(* CODESYS project lc.library
   DefaultNamespace: KOSTAL.AF2024.Connectivity.LC
   DocFormat: reStructuredText
   Description: Contains Components to communicate with LC Webservice.
      
      Designed with webAPI Version 2.0.39
      
      =====================
      BASED NOT ON I_LC!!
      =====================
   Author: Frank Dümpelmann
   Title: KOSTAL.AF2024.Connectivity.LC
   Version: 1.0.0.0
   Company: KOSTAL GmbH & Co.KG
   Placeholder: KOSTAL.AF2024.Connectivity.LC

Project tree, tasks and I/O mapping:
  libraries: KOSTAL.AF2024.Connectivity.TLS.CipherSuite.OpenSSL, 1.0.0.0 (KOSTAL GmbH & Co.KG); KOSTAL.AF2024.Core.FileLogger, 1.0.0.0 (KOSTAL GmbH & Co.KG); KOSTAL.AF2024.Core.functionResponse, 1.0.0.0 (KOSTAL GmbH & Co.KG); KOSTAL.AF2024.Core.GetSystemTime, 1.0.1.0 (KOSTAL GmbH & Co.KG); KOSTAL.AF2024.Core.JsonTools, 1.0.0.0 (KOSTAL GmbH & Co.KG); KOSTAL.AF2024.Core.ListOf, 1.0.0.0 (KOSTAL GmbH & Co.KG); KOSTAL.AF2024.Core.Process, 1.0.1.0 (KOSTAL GmbH & Co.KG); KOSTAL.AF2024.Core.Settings, 1.0.0.0 (KOSTAL GmbH & Co.KG); KOSTAL.AF2024.Core.StringTools, 1.0.0.0 (KOSTAL GmbH & Co.KG); KOSTAL.AF2024.Core.System, 1.0.0.0 (KOSTAL GmbH & Co.KG); Tc2_Standard, 3.4.5.0 (Beckhoff Automation GmbH); Tc2_System, 3.6.4.0 (Beckhoff Automation GmbH); Tc2_Utilities, 3.7.4.0 (Beckhoff Automation GmbH); Tc3_IotBase, 3.4.5.0 (Beckhoff Automation GmbH); Tc3_JsonXml, 3.4.4.0 (Beckhoff Automation GmbH)
  0_Internal/
    interface _I_T_Copy: CopyTo
    interface _I_T_Copy_Owner: Clear, CopyFrom, CopyTo
    interface _I_T_CopyFrom: CopyFrom
    function block _T_Copy [ST]: Clear, CopyFrom, CopyTo
  1_Config/
    Reader/
      DUT/
        interface I_T_Header: CopyTo, ID, name, sourceName, timeStamp
        interface I_T_Header_CopyFrom: CopyFrom
        function block T_Header [ST]: Clear, CopyFrom, CopyTo, ID, name, sourceName, timeStamp
      function block FB_Reader [ST]: _Step_ClearContent, _Step_ParseContent, CFG, Header
      global variables JSON_MEMBER
    interface I_T_CFG: ClientName, ClientProcess, CopyTo, HostName, HostPort, Valid
    interface I_T_CFG_CopyFrom: CopyFrom
    function block T_CFG [ST]: Clear, ClientName, ClientProcess, CopyFrom, CopyTo, HostName, HostPort, Valid
  2_BaseClass/
    DUT/
      Response/
        interface I_T_ResponseResult: CopyTo, errorMessage, internalDuration, isErrorOccured, isResultGood
        interface I_T_ResponseResult_CopyFrom: CopyFrom
        interface I_T_ResponseResult_Owner: clear, CopyFrom, CopyTo, errorMessage, internalDuration, isErrorOccured, isResultGood
        function block T_ResponseResult [ST]: clear, CopyFrom, CopyTo, errorMessage, internalDuration, isErrorOccured, isResultGood
      data type E_PROCESS
      data type E_Verbose
    POE/
      function block FB_LC [ST]: _getResponseResultFromJson, _PARSE_ARRAY, _PARSE_BOOL, _PARSE_BYTE, _PARSE_DINT, _PARSE_JSON, _PARSE_STRING, _PARSE_TIME, _PARSE_UDINT, _PARSE_ULINT, _00_clientCfg, _01_Ready, _10_finishFail, _10_finishPass, _10_GET, _10_GET_CTRL, _10_GET_ResponseResult, _10_GET_ResponseResult_CTRL, _10_SET, _10_SET_CTRL, _99_stepError, _CfgChange, _CfgHasChanged, _deviceDefine, _logStartMessage, _UriGet, _UrlReplace, _VerboseHandler, ClientName, ClientProcess, HostName, HostPort, HTTP_Statuscode, IN_PROCESS, KeepAlive, repeatsOnFail, State, TimeOut, WS_Duration, FBmain, GetTimeStamp, linkConfig, LinkTime, RedirectClient, Verbose, _FBmain
  3_DUT/
    OptionalFlags/
      interface I_T_OptionalFlags: FlagsInRange, get
      interface I_T_OptionalFlags_Owner: clear, FlagsInRange, get, set
      function block T_OptionalFlags [ST]: clear, CopyFrom, FlagsInRange, get, set
    OptionalStrings/
      interface I_T_OptionalStrings: get, StringsInRange
      interface I_T_OptionalStrings_Owner: clear, get, set, StringsInRange
      function block T_OptionalStrings [ST]: clear, CopyFrom, get, set, StringsInRange
    PreviousProcess/
      ListOf/
        function block FB_ListOfPreviousProcess [ST]: _get_I, _get_I_Owner, _removePayLoad, _verifyMember, Add_DUT, Clear, CopyFrom, CopyTo, Delete_DUT, Get_I, Get_I_ByProcessName, Get_I_Owner, NumberOfMember
        interface I_ListOfPreviousProcess: CopyTo, Get_I, Get_I_ByProcessName, NumberOfMember
        interface I_ListOfPreviousProcess_CopyFrom: CopyFrom
        interface I_ListOfPreviousProcess_Owner: Add_DUT, Clear, CopyFrom, CopyTo, Delete_DUT, Get_I, Get_I_ByProcessName, Get_I_Owner, NumberOfMember
      interface I_T_PreviousProcess: articlenumberRegex, databaseName, PreviousProcesses, processName, processStamp, searchMode, useOnlyTable
      interface I_T_PreviousProcess_Owner: articlenumberRegex, clear, databaseName, PreviousProcesses_Owner, processName, processStamp, searchMode, useOnlyTable
      function block T_PreviousProcess [ST]: articlenumberRegex, clear, CopyFrom, databaseName, PreviousProcesses, PreviousProcesses_Owner, processName, processStamp, searchMode, useOnlyTable
    ProcessConfig/
      ListOf/
        function block FB_ListOfProcessConfig [ST]: _get_I, _get_I_Owner, _removePayLoad, _verifyMember, Add_DUT, Clear, CopyFrom, CopyTo, Delete_DUT, Get_I, Get_I_Owner, NumberOfMember
        interface I_ListOfProcessConfig: CopyTo, Get_I, NumberOfMember
        interface I_ListOfProcessConfig_CopyFrom: CopyFrom
        interface I_ListOfProcessConfig_Owner: Add_DUT, Clear, CopyFrom, CopyTo, Delete_DUT, Get_I, Get_I_Owner, NumberOfMember
      interface I_T_ProcessConfig: activeCheckFQDN, allowedFQDN, articlenumberRegex, PreviousProcesses, serialnumberRegex, traceID
      interface I_T_ProcessConfig_Owner: activeCheckFQDN, allowedFQDN, articlenumberRegex, clear, PreviousProcesses_Owner, serialnumberRegex, traceID
      function block T_ProcessConfig [ST]: activeCheckFQDN, allowedFQDN, articlenumberRegex, clear, CopyFrom, PreviousProcesses, PreviousProcesses_Owner, serialnumberRegex, traceID
    SingleProcess/
      ListOf/
        function block FB_ListOfSingleProcess [ST]: _get_I, _get_I_Owner, _removePayLoad, _verifyMember, Add_DUT, Clear, CopyFrom, CopyTo, Delete_DUT, Get_I, Get_I_Owner, NumberOfMember
        interface I_ListOfSingleProcess: CopyTo, Get_I, NumberOfMember
        interface I_ListOfSingleProcess_CopyFrom: CopyFrom
        interface I_ListOfSingleProcess_Owner: Add_DUT, Clear, CopyFrom, CopyTo, Delete_DUT, Get_I, Get_I_Owner, NumberOfMember
      interface I_T_SingleProcess: articleNumber, id, OptionalFlags, OptionalStrings, process, result, serialNumber, timeStamp, traceId
      interface I_T_SingleProcess_Owner: articleNumber, clear, id, OptionalFlags_Owner, OptionalStrings_Owner, process, result, serialNumber, timeStamp, traceId
      function block T_SingleProcess [ST]: articleNumber, clear, CopyFrom, id, OptionalFlags, OptionalFlags_Owner, OptionalStrings, OptionalStrings_Owner, process, result, serialNumber, timeStamp, traceId
    SubModule/
      ListOf/
        function block FB_ListOfSubModule [ST]: _get_I, _get_I_Owner, _removePayLoad, _verifyMember, Add_DUT, Clear, CopyFrom, CopyTo, Delete_DUT, Get_I, Get_I_Owner, NumberOfMember
        interface I_ListOfSubModule: CopyTo, Get_I, NumberOfMember
        interface I_ListOfSubModule_CopyFrom: CopyFrom
        interface I_ListOfSubModule_Owner: Add_DUT, Clear, CopyFrom, CopyTo, Delete_DUT, Get_I, Get_I_Owner, NumberOfMember
      interface I_T_SubModule: articleNumber, serialNumber
      interface I_T_SubModule_Owner: articleNumber, clear, serialNumber
      function block T_SubModule [ST]: articleNumber, clear, CopyFrom, serialNumber
    SubModuleOfProcess/
      ListOf/
        function block FB_ListOfSubModuleOfProcess [ST]: _get_I, _get_I_Owner, _removePayLoad, _verifyMember, Add_DUT, Clear, CopyFrom, CopyTo, Delete_DUT, Get_I, Get_I_Owner, NumberOfMember
        interface I_ListOfSubModuleOfProcess: CopyTo, Get_I, NumberOfMember
        interface I_ListOfSubModuleOfProcess_CopyFrom: CopyFrom
        interface I_ListOfSubModuleOfProcess_Owner: Add_DUT, Clear, CopyFrom, CopyTo, Delete_DUT, Get_I, Get_I_Owner, NumberOfMember
      interface I_T_SubModuleOfProcess: timeStamp
      interface I_T_SubModuleOfProcess_Owner: timeStamp
      function block T_SubModuleOfProcess [ST]: clear, CopyFrom, timeStamp
    WriteCurrentStampDataDto/
      interface I_T_WriteCurrentStampDataDto: articleNumber, OptionalFlags, OptionalStrings, result, serialNumber
      interface I_T_WriteCurrentStampDataDto_Owner: articleNumber, clear, OptionalFlags_Owner, OptionalStrings_Owner, result, serialNumber
      function block T_WriteCurrentStampDataDto [ST]: articleNumber, clear, CopyFrom, OptionalFlags, OptionalFlags_Owner, OptionalStrings, OptionalStrings_Owner, result, serialNumber
  4_GVL/
    global variables API_VERSION
    global variables PROCESS_CONFIG
    global variables PROCESS_INFO
    global variables RESPONSE_BODY
    global variables SETTINGS
    global variables SUBMODUL_INFO
    global variables URL
  5_POU/
    GetetParentBySubmoduleSerialnumber/
      function block FB_GetParent_By_SM_SN [ST]: _getProcessInfo, _getSubModule_n, _getSubModuleList, _01_Ready, _10_getProcessInfo, _10_getSubModule_n, _10_getSubModuleList, _10_processRead, _selectUrl, Execute, ListOfSubModules, ResponseProcess, ResponseResult, _FBmain
    GetSubModulesByParentSerialNumber/
      function block FB_GetSM_ByParentSN [ST]: _getProcessInfo, _getSubModule_n, _getSubModuleList, _01_Ready, _10_getProcessInfo, _10_getSubModule_n, _10_getSubModuleList, _10_processRead, _selectUrl, Execute, ListOfSubModules, ResponseProcess, ResponseResult, _FBmain
    Init/
      function block FB_Init [ST]
    ReadApiVersion/
      MustBeExtended/
        function block _FB_ReadApiVersion [ST]: _getApiVersion, _01_Ready, _10_getapiVersion, _10_processRead, _selectUrl, apiVersion, ResponseResult, _FBmain
      function block FB_ReadApiVersion [ST]: Execute, _selectUrl
    ReadProcess/
      MustBeExtended/
        function block _FB_ReadProcess [ST]: _getProcessInfo, _getProcessInfoList, _01_Ready, _10_getProcessInfo_n, _10_getProcessInfoList, _10_processRead, _selectUrl, GetSingleProcess, NumberOfSingleProcess, ProcessInfoListLenght, ResponseResult, _FBmain
      function block FB_ReadPreviousProcess_SN [ST]: Execute, _selectUrl
      function block FB_ReadPreviousProcess_SN_ART [ST]: Execute, _selectUrl
      function block FB_ReadProcess_ID [ST]: Execute, _selectUrl
      function block FB_ReadProcess_SN [ST]: Execute, _selectUrl
      function block FB_ReadProcess_SN_ART [ST]: Execute, _selectUrl
    ReadProcessConfig/
      MustBeExtended/
        function block _FB_ReadConfig [ST]: _getPreviousProcess, _getPreviousProcesses, _getPreviousProcessList, _getProcessConfig, _getProcessConfigList, _01_Ready, _10_getProcessConfig_n, _10_getProcessConfigList, _10_processRead, _selectUrl, GetProcessConfig, NumberOfProcessConfig, ResponseResult, _FBmain
      function block FB_ReadProcessConfig [ST]: Execute, _selectUrl
    WriteProcess/
      MustBeExtended/
        function block _FB_WriteProcess [ST]: _getProcessInfo, _01_Ready, _10_getProcessInfo, _10_processWrite, _20_setProcessInfo, _selectUrl, Execute, ResponseProcess, ResponseResult, WriteDataDto
      function block FB_WriteProcess [ST]: _selectUrl, _FBmain
      function block FB_WriteProcessWithSM [ST]: _20_setSubModules, _selectUrl, ListOfSubModules, _FBmain
  Project Information/
    function F_GetCompany [ST]
    function F_GetTitle [ST]
    function F_GetVersion [ST]
  Version/
    global variables Global_Version
*)

// 2_BaseClass/DUT/E_PROCESS
{attribute 'qualified_only'}
{attribute 'strict'}
TYPE E_PROCESS :
(
	idle		:= 0,
	execute	:= 1
);
END_TYPE

// 2_BaseClass/DUT/E_Verbose
{attribute 'qualified_only'}
{attribute 'strict'}
(*
Note that the verbose status is evaluated binary
================================================
*)
TYPE E_Verbose :
(
	none 			:= 0,
	Request		:= 1,
	Response	:= 2,
	Both			:= 3
);
END_TYPE

// 1_Config/Reader/JSON_MEMBER
{attribute 'qualified_only'}
VAR_GLOBAL CONSTANT

	{region 'Header'}
		ID					: STRING:= 'ID';
		name				: STRING:= 'name'; 
		timeStamp		: STRING:= 'timeStamp'; 
		sourceName	: STRING:= 'sourceName'; 
	{endregion}

	{region 'LC'}
		LC						: STRING:= 'LC';
		HostName			: STRING:= 'HostName';
		HostPort			: STRING:= 'HostPort';
		ClientName		: STRING:= 'ClientName';
		ClientProcess	: STRING:= 'ClientProcess';
	{endregion}

END_VAR

// 4_GVL/API_VERSION
{attribute 'qualified_only'}
VAR_GLOBAL
	apiVersion		:	STRING:= 'apiVersion';
END_VAR

// 4_GVL/PROCESS_CONFIG
{attribute 'qualified_only'}
VAR_GLOBAL CONSTANT
	//
	processConfiguration	:	STRING:=	'processConfiguration';
	//
  articlenumberRegex	: STRING:=	'articlenumberRegex';	//"^[0-9]{8}-(([0-9]{2})|([0-9]{4}))$",
  serialnumberRegex		: STRING:=	'serialnumberRegex';	//"^([A-Z0-9]{13})$|^([0-9]{14})$",
  traceID							: STRING:=	'traceID';	//99056,
	activeCheckFQDN			: STRING:=	'activeCheckFQDN';
	allowedFQDN					: STRING:=	'allowedFQDN';
	///--
  previousProcesses	: STRING:=	'previousProcesses';	//[...]
	//
  processName			: STRING:=	'processName';	//"ASS01",
  processStamp		: STRING:=	'processStamp';	//"ASS01",
  databaseName		: STRING:=	'databaseName';		//"test",
  useOnlyTable		: STRING:=	'useOnlyTable';	//"lc_test"
  searchMode			: STRING:=	'searchMode';	//0,
  //articlenumberRegex	: STRING:=	'articlenumberRegex';	same as in parent node
  //previousProcesses	: STRING:=	'previousProcesses';	same as in parent node

//obsolete
//  databaseServer	:	STRING:=	'databaseServer';	//"debelc034.de.kostal.int",
//  databasePort		: STRING:=	'databasePort';		//3306,
//  databaseUser		: STRING:=	'databaseUser';		//null,
END_VAR

// 4_GVL/PROCESS_INFO
{attribute 'qualified_only'}
VAR_GLOBAL CONSTANT
	//
	processInfoList	: STRING:= 'processInfoList'; 
	processInfo			: STRING:= 'processInfo';
	//
	id								: STRING:= 'id';
	serialNumber			: STRING:= 'serialNumber';
	articleNumber			: STRING:= 'articleNumber';
	timeStamp					: STRING:= 'timeStamp';
	traceId						: STRING:= 'traceId';
	process						: STRING:= 'process';
	result						: STRING:= 'result';
	optionalString_1	: STRING:= 'optionalString_1';
	optionalString_2	: STRING:= 'optionalString_2';
	optionalString_3	: STRING:= 'optionalString_3';
	optionalString_4	: STRING:= 'optionalString_4';
	optionalFlag_1		: STRING:= 'optionalFlag_1';
	optionalFlag_2		: STRING:= 'optionalFlag_2';
	optionalFlag_3		: STRING:= 'optionalFlag_3';
	optionalFlag_4		: STRING:= 'optionalFlag_4';
	optionalFlag_5		: STRING:= 'optionalFlag_5';
	optionalFlag_6		: STRING:= 'optionalFlag_6';
	optionalFlag_7		: STRING:= 'optionalFlag_7';
	optionalFlag_8		: STRING:= 'optionalFlag_8';

	//
	childs	: STRING:= 'Childs';
																		
END_VAR

// 4_GVL/RESPONSE_BODY
{attribute 'qualified_only'}
VAR_GLOBAL CONSTANT
	
	isErrorOccured		:	STRING:= 'isErrorOccured';
	isResultGood			:	STRING:= 'isResultGood';
	errorMessage			:	STRING:= 'errorMessage';
	internalDuration	:	STRING:= 'internalDuration';
	
END_VAR

// 4_GVL/SETTINGS
{attribute 'qualified_only'}
VAR_GLOBAL CONSTANT
	OPTIONAL_FLAGS_MAX				: UINT:= 8;
	
	OPTIONAL_STRINGS_MAX			: UINT:= 4;
	OPTIONAL_STRINGS_LENGHT		: UINT:= SIZEOF(KOSTAL_AF2024_Core_Settings.T_MaxString_UTF8);
END_VAR

// 4_GVL/SUBMODUL_INFO
{attribute 'qualified_only'}
VAR_GLOBAL CONSTANT
	//
	subModules	: STRING:= 'submodules';
	//
	serialNumber	: STRING:=	'serialNumber';
	articleNumber : STRING:=	'articleNumber';
	timestamp			: STRING:=	'timestamp';	//only in S´sub modules of process available
END_VAR

// 4_GVL/URL
{attribute 'qualified_only'}
VAR_GLOBAL CONSTANT

	URI_BASE	: KOSTAL_AF2024_Core_Settings.T_MaxString_UTF8:=  '/ws/api/gen2/';
	
	READ_API_VERSION	: KOSTAL_AF2024_Core_Settings.T_MaxString_UTF8:= 'readApiVersion';
	
	READ_PROC_RECORD_ID	: KOSTAL_AF2024_Core_Settings.T_MaxString_UTF8:= 'readProcess/{ClientName}/{ClientProcess}/id={RecordID}';

	READ_PROC_SERNO				: KOSTAL_AF2024_Core_Settings.T_MaxString_UTF8:= 'readProcess/{ClientName}/{ClientProcess}/{SerialNumber}';
	READ_PROCESS_SERNO_OPT_PROC	: KOSTAL_AF2024_Core_Settings.T_MaxString_UTF8:= 'readProcess/{ClientName}/{ClientProcess}/{SerialNumber}?Process={?Process=}';
	
	READ_PROC_SERNO_ARTNO			: KOSTAL_AF2024_Core_Settings.T_MaxString_UTF8:= 'readProcess/{ClientName}/{ClientProcess}/{SerialNumber}/{ArticleNumber}';
	READ_PROC_SERNO_ARTNO_OPT_PROC	: KOSTAL_AF2024_Core_Settings.T_MaxString_UTF8:= 'readProcess/{ClientName}/{ClientProcess}/{SerialNumber}/{ArticleNumber}?Process={?Process=}';

	READ_PREV_PROC_SERNO	: KOSTAL_AF2024_Core_Settings.T_MaxString_UTF8:= 'readPreviousProcess/{ClientName}/{ClientProcess}/{SerialNumber}';

	READ_PREV_PROC_SERNO_ARTNO	: KOSTAL_AF2024_Core_Settings.T_MaxString_UTF8:= 'readPreviousProcess/{ClientName}/{ClientProcess}/{SerialNumber}/{ArticleNumber}';
	
	WRITE_CUR_PROC					: KOSTAL_AF2024_Core_Settings.T_MaxString_UTF8:= 'writeCurrentProcess/{ClientName}/{ClientProcess}';
	WRITE_CUR_PROC_WITH_SUBMODULS	: KOSTAL_AF2024_Core_Settings.T_MaxString_UTF8:= 'writeCurrentProcessWithSubmodules/{ClientName}/{ClientProcess}';

	READ_PROC_CONF			: KOSTAL_AF2024_Core_Settings.T_MaxString_UTF8:= 'readProcessConfig/{ClientName}';
	READ_PROC_CONF_OPT_PROC	: KOSTAL_AF2024_Core_Settings.T_MaxString_UTF8:= 'readProcessConfig/{ClientName}/{ClientProcess}';

	READ_SUB_MODULES_BY_PARENT_SERIAL_NUMBER	: KOSTAL_AF2024_Core_Settings.T_MaxString_UTF8:= 'getSubmodulesByParentserialnumber/{ClientName}/{ClientProcess}/{ParentSerialnumber}';
	READ_PARENT_BY_SUB_MODULE_SERIAL_NUMBER		: KOSTAL_AF2024_Core_Settings.T_MaxString_UTF8:= 'getParentBySubmoduleSerialnumber/{ClientName}/{ClientProcess}/{SubmoduleSerialnumber}';
END_VAR

//Placeholder for URI
{attribute 'qualified_only'}
VAR_GLOBAL CONSTANT
	PLACEHOLDER_CLIENT_NAME						: STRING:= '{ClientName}';
	PLACEHOLDER_CLIENT_PROCESS				: STRING:= '{ClientProcess}';
	PLACEHOLDER_RECORD_ID							: STRING:= '{RecordID}';
	PLACEHOLDER_SERIALNUMBER					: STRING:= '{SerialNumber}';
	PLACEHOLDER_ARTICLENUMBER					: STRING:= '{ArticleNumber}';
	PLACEHOLDER_OPTIONAL_PROCESS			: STRING:= '{?Process=}';

	PLACEHOLDER_PARENT_SERIAL_NUMBER	: STRING:= '{ParentSerialnumber}';
	PLACEHOLDER_SUB_MODULE_SERIAL_NUMBER		: STRING:= '{SubmoduleSerialnumber}';
END_VAR

// Version/Global_Version
{attribute 'TcGenerated'}
{attribute 'no-analysis'}
{attribute 'linkalways'}
// This function has been automatically generated from the project information.
VAR_GLOBAL CONSTANT
	{attribute 'const_non_replaced'}
	stLibVersion_KOSTAL_AF2024_Connectivity_LC : ST_LibVersion := (iMajor := 1, iMinor := 0, iBuild := 0, iRevision := 0, nFlags := 1, sVersion := '1.0.0.0');
END_VAR

// 0_Internal/_I_T_Copy
INTERFACE _I_T_Copy EXTENDS KOSTAL_AF2024_Core_System.I_Interface

METHOD PUBLIC CopyTo : BOOL
VAR_INPUT
	IN	: KOSTAL_AF2024_Core_System.I_Interface;
END_VAR
END_METHOD

END_INTERFACE

// 0_Internal/_I_T_Copy_Owner
INTERFACE _I_T_Copy_Owner EXTENDS KOSTAL_AF2024_Core_System.I_Interface

METHOD PUBLIC Clear
END_METHOD

METHOD PUBLIC CopyFrom : BOOL
VAR_INPUT
	IN	: KOSTAL_AF2024_Core_System.I_Interface;
END_VAR
END_METHOD

METHOD PUBLIC CopyTo : BOOL
VAR_INPUT
	IN	: KOSTAL_AF2024_Core_System.I_Interface;
END_VAR
END_METHOD

END_INTERFACE

// 0_Internal/_I_T_CopyFrom
INTERFACE _I_T_CopyFrom EXTENDS KOSTAL_AF2024_Core_System.I_Interface

METHOD PUBLIC CopyFrom : BOOL
VAR_INPUT
	IN	: KOSTAL_AF2024_Core_System.I_Interface;
END_VAR
END_METHOD

END_INTERFACE

// 0_Internal/_T_Copy
FUNCTION_BLOCK ABSTRACT _T_Copy IMPLEMENTS _I_T_Copy, _I_T_Copy_Owner, _I_T_CopyFrom

METHOD PUBLIC Clear
END_METHOD

METHOD PUBLIC CopyFrom : BOOL
VAR_INPUT
	IN	: KOSTAL_AF2024_Core_System.I_Interface;
END_VAR

VAR
	_IN	: KOSTAL_AF2024_Core_System.I_Interface;
END_VAR


CopyFrom:= (IN <> 0) AND_THEN __QUERYINTERFACE(IN, _IN) AND_THEN (_IN <> 0);
END_METHOD

METHOD PUBLIC CopyTo : BOOL
VAR_INPUT
	IN	: KOSTAL_AF2024_Core_System.I_Interface;
END_VAR

VAR
	_IN	: _I_T_CopyFrom;
END_VAR

IF (IN = 0) OR_ELSE NOT __QUERYINTERFACE(IN, _IN) OR_ELSE (_IN = 0) THEN	RETURN;	END_IF

CopyTo:= _IN.CopyFrom(THIS^);
END_METHOD

END_FUNCTION_BLOCK

// 1_Config/Reader/DUT/I_T_Header
INTERFACE I_T_Header EXTENDS KOSTAL_AF2024_Core_System.I_Interface

METHOD PUBLIC CopyTo : BOOL
VAR_INPUT
	IN	: I_T_Header_CopyFrom;
END_VAR
END_METHOD

PROPERTY PUBLIC ID : KOSTAL_AF2024_Core_Settings.T_MaxString_UTF8
GET
END_GET
END_PROPERTY

PROPERTY PUBLIC name : KOSTAL_AF2024_Core_Settings.T_MaxString_UTF8
GET
END_GET
END_PROPERTY

PROPERTY PUBLIC sourceName : KOSTAL_AF2024_Core_Settings.T_MaxString_UTF8
GET
END_GET
END_PROPERTY

PROPERTY PUBLIC timeStamp : KOSTAL_AF2024_Core_Settings.T_MaxString_UTF8
GET
END_GET
END_PROPERTY

END_INTERFACE

// 1_Config/Reader/DUT/I_T_Header_CopyFrom
INTERFACE I_T_Header_CopyFrom EXTENDS KOSTAL_AF2024_Core_System.I_Interface

METHOD PUBLIC CopyFrom
VAR_INPUT
	IN	: KOSTAL_AF2024_Core_System.I_Interface;
END_VAR
END_METHOD

END_INTERFACE

// 1_Config/Reader/DUT/T_Header
FUNCTION_BLOCK PUBLIC T_Header IMPLEMENTS I_T_Header, I_T_Header_CopyFrom

VAR
	_ID					: KOSTAL_AF2024_Core_Settings.T_MaxString_UTF8;
	_name				: KOSTAL_AF2024_Core_Settings.T_MaxString_UTF8;
	_timeStamp	: KOSTAL_AF2024_Core_Settings.T_MaxString_UTF8;
	_sourceName	: KOSTAL_AF2024_Core_Settings.T_MaxString_UTF8;	
END_VAR

METHOD PUBLIC Clear
VAR_INPUT
END_VAR

_ID					:= '';
_name				:= '';
_sourceName	:= '';
_timeStamp	:= '';
END_METHOD

METHOD PUBLIC CopyFrom
VAR_INPUT
	IN	: KOSTAL_AF2024_Core_System.I_Interface;
END_VAR

VAR
	_IN	: I_T_Header;
END_VAR

IF IN = 0 THEN	RETURN;	END_IF
IF NOT __QUERYINTERFACE(IN, _IN) OR_ELSE _IN = 0 THEN RETURN;	END_IF

_ID					:= _IN.ID;
_name				:= _IN.name;
_timeStamp	:= _IN.timeStamp;
_sourceName	:= _IN.sourceName;
END_METHOD

METHOD PUBLIC CopyTo : BOOL
VAR_INPUT
	IN	: I_T_Header_CopyFrom;
END_VAR

IF IN = 0 THEN	RETURN;	END_IF

IN.CopyFrom(THIS^);
END_METHOD

PROPERTY PUBLIC ID : KOSTAL_AF2024_Core_Settings.T_MaxString_UTF8
GET

ID:= _ID;
END_GET
SET

_ID:= ID;
END_SET
END_PROPERTY

PROPERTY PUBLIC name : KOSTAL_AF2024_Core_Settings.T_MaxString_UTF8
GET

name:= _name;
END_GET
SET

_name:= name;
END_SET
END_PROPERTY

PROPERTY PUBLIC sourceName : KOSTAL_AF2024_Core_Settings.T_MaxString_UTF8
GET

sourceName:= _sourceName;
END_GET
SET

_sourceName:= sourceName;
END_SET
END_PROPERTY

PROPERTY PUBLIC timeStamp : KOSTAL_AF2024_Core_Settings.T_MaxString_UTF8
GET

timeStamp:= _timeStamp;
END_GET
SET

_timeStamp:= timeStamp;
END_SET
END_PROPERTY

END_FUNCTION_BLOCK

// 1_Config/Reader/FB_Reader
FUNCTION_BLOCK PUBLIC FB_Reader EXTENDS KOSTAL_AF2024_Core_JsonTools._FB_Base_RO
VAR
	_Header	: T_Header;
	_CFG		: T_CFG;
END_VAR

METHOD PROTECTED _Step_ClearContent
VAR_INPUT
END_VAR

_Header.Clear();
_CFG.Clear();

SUPER^._Step_ClearContent();
END_METHOD

METHOD PROTECTED _Step_ParseContent
VAR_INPUT
END_VAR

VAR
	_key		: KOSTAL_AF2024_Core_Settings.T_MaxString_UTF8;
	_value	: KOSTAL_AF2024_Core_Settings.T_MaxString_UTF8;
	_resp		: KOSTAL_AF2024_Core_Settings.T_MaxString_UTF8;
	_jLC		: Tc3_IotBase.SJsonValue;
END_VAR
//===================================================================================
//Header
//===================================================================================
_key:= JSON_MEMBER.ID;
_Header.ID:= _PARSE_STRING(_jDoc, _key, TRUE, _resp);

IF _resp <> '' THEN
	_State.description:= Tc2_Standard.WCONCAT(TO_WSTRING(_resp), "; ID is empty > not allowed");
	_step.set(_ADDRESS_FINISH_FAIL);
	RETURN;
END_IF


//===================================================================================
_key:= JSON_MEMBER.name;
_Header.name:= _PARSE_STRING(_jDoc, _key, FALSE, 0);

//===================================================================================
_key:= JSON_MEMBER.timeStamp;
_Header.timeStamp:= _PARSE_STRING(_jDoc, _key, FALSE, 0);

//===================================================================================
_key:= JSON_MEMBER.sourceName;
_Header.sourceName:= _PARSE_STRING(_jDoc, _key, FALSE, 0);


//===================================================================================
//LC
//===================================================================================
_key:= JSON_MEMBER.LC;
_jLC:= _PARSE_JSON(_jDoc, _key, TRUE, _resp);
 
IF _resp <> '' THEN
	_State.description:= Tc2_Standard.WCONCAT(TO_WSTRING(_resp), "; LC nnode is empty > not allowed");
	_step.set(_ADDRESS_FINISH_FAIL);
	RETURN;
END_IF

IF _jLC = 0 THEN
	_State.description:= "LC nnode does not exist > not allowed";
	_step.set(_ADDRESS_FINISH_FAIL);
	RETURN;
END_IF

//===================================================================================
_key:= JSON_MEMBER.HostName;
_CFG.HostName:= _PARSE_STRING(_jLC, _key, TRUE, _resp);

IF _resp <> '' THEN
	_State.description:= Tc2_Standard.WCONCAT(TO_WSTRING(_resp), "; Hostname failed > not allowed");
	_step.set(_ADDRESS_FINISH_FAIL);
	RETURN;
END_IF

IF _CFG.HostName = '' THEN
	_State.description:= "Hostname is empty > not allowed";
	_step.set(_ADDRESS_FINISH_FAIL);
	RETURN;
END_IF

//===================================================================================
_key:= JSON_MEMBER.HostPort;
_CFG.HostPort:= UDINT_TO_UINT(_PARSE_UDINT(_jLC, _key, FALSE, 0));

//===================================================================================
_key:= JSON_MEMBER.ClientName;
_CFG.ClientName:= _PARSE_STRING(_jLC, _key, TRUE, _resp);

IF _resp <> '' THEN
	_State.description:= Tc2_Standard.WCONCAT(TO_WSTRING(_resp), "; Clientname failed > not allowed");
	_step.set(_ADDRESS_FINISH_FAIL);
	RETURN;
END_IF

IF _CFG.ClientName = '' THEN
	_State.description:= "ClientName is empty > not allowed";
	_step.set(_ADDRESS_FINISH_FAIL);
	RETURN;
END_IF

//===================================================================================
_key:= JSON_MEMBER.ClientProcess;
_CFG.ClientProcess:= _PARSE_STRING(_jLC, _key, TRUE, _resp);

IF _resp <> '' THEN
	_State.description:= Tc2_Standard.WCONCAT(TO_WSTRING(_resp), "; ClientProcess failed > not allowed");
	_step.set(_ADDRESS_FINISH_FAIL);
	RETURN;
END_IF

IF _CFG.ClientProcess = '' THEN
	_State.description:= "ClientProcess is empty > not allowed";
	_step.set(_ADDRESS_FINISH_FAIL);
	RETURN;
END_IF

//===================================================================================
_CFG.Valid:= TRUE;

SUPER^._Step_ParseContent();
END_METHOD

PROPERTY PUBLIC CFG :I_T_CFG
GET

CFG:= _CFG;
END_GET
END_PROPERTY

PROPERTY PUBLIC Header : I_T_Header
GET

Header:= _Header;
END_GET
END_PROPERTY

END_FUNCTION_BLOCK

// 1_Config/T_CFG
FUNCTION_BLOCK PUBLIC T_CFG IMPLEMENTS I_T_CFG, I_T_CFG_CopyFrom

VAR
	_HostName				:	KOSTAL_AF2024_Core_Settings.T_MaxString_UTF8;
	_HostPort				: UINT;
	_ClientName			: KOSTAL_AF2024_Core_Settings.T_MaxString_UTF8;
	_ClientProcess	: KOSTAL_AF2024_Core_Settings.T_MaxString_UTF8;
	_Valid					: BOOL;	//set contains valid data 
END_VAR

METHOD PUBLIC Clear

_HostName				:= '';
_HostPort				:= UINT#0;
_ClientName			:= '';
_ClientProcess	:= '';
_Valid					:= FALSE;
END_METHOD

PROPERTY PUBLIC ClientName : KOSTAL_AF2024_Core_Settings.T_MaxString_UTF8
GET

ClientName:= _ClientName;
END_GET
SET

_ClientName:= ClientName;
END_SET
END_PROPERTY

PROPERTY PUBLIC ClientProcess : KOSTAL_AF2024_Core_Settings.T_MaxString_UTF8
GET

ClientProcess:= _ClientProcess;
END_GET
SET

_ClientProcess:= ClientProcess;
END_SET
END_PROPERTY

METHOD PUBLIC CopyFrom
VAR_INPUT
	IN	: KOSTAL_AF2024_Core_System.I_Interface;
END_VAR

VAR
	_IN	: I_T_CFG;
END_VAR

IF IN = 0 THEN	RETURN;	END_IF
IF NOT __QUERYINTERFACE(IN, _IN) OR_ELSE _IN= 0 THEN RETURN;	END_IF

_HostName				:= _IN.HostName;
_HostPort				:= _IN.HostPort;
_ClientName			:= _IN.ClientName;
_ClientProcess	:= _IN.ClientProcess;
_Valid					:= _IN.Valid;
END_METHOD

METHOD PUBLIC CopyTo
VAR_INPUT
	IN	: I_T_CFG_CopyFrom;
END_VAR

IF IN = 0 THEN	RETURN;	END_IF

IN.CopyFrom(THIS^);
END_METHOD

PROPERTY PUBLIC HostName : KOSTAL_AF2024_Core_Settings.T_MaxString_UTF8
GET

HostName:= _HostName;
END_GET
SET

_HostName:= HostName;
END_SET
END_PROPERTY

PROPERTY PUBLIC HostPort : UINT
GET

HostPort:= _HostPort;
END_GET
SET

_HostPort:= HostPort;
END_SET
END_PROPERTY

PROPERTY PUBLIC Valid : BOOL
GET

Valid:= _Valid;
END_GET
SET

_Valid:= Valid;
END_SET
END_PROPERTY

END_FUNCTION_BLOCK

// 1_Config/I_T_CFG
INTERFACE I_T_CFG EXTENDS KOSTAL_AF2024_Core_System.I_Interface

PROPERTY PUBLIC ClientName : KOSTAL_AF2024_Core_Settings.T_MaxString_UTF8
GET
END_GET
END_PROPERTY

PROPERTY PUBLIC ClientProcess : KOSTAL_AF2024_Core_Settings.T_MaxString_UTF8
GET
END_GET
END_PROPERTY

METHOD PUBLIC CopyTo
VAR_INPUT
	IN	: I_T_CFG_CopyFrom;
END_VAR
END_METHOD

PROPERTY PUBLIC HostName : KOSTAL_AF2024_Core_Settings.T_MaxString_UTF8
GET
END_GET
END_PROPERTY

PROPERTY PUBLIC HostPort : UINT
GET
END_GET
END_PROPERTY

PROPERTY PUBLIC Valid : BOOL
GET
END_GET
END_PROPERTY

END_INTERFACE

// 1_Config/I_T_CFG_CopyFrom
INTERFACE I_T_CFG_CopyFrom EXTENDS KOSTAL_AF2024_Core_System.I_Interface

METHOD PUBLIC CopyFrom
VAR_INPUT
	IN	: KOSTAL_AF2024_Core_System.I_Interface;
END_VAR
END_METHOD

END_INTERFACE

// 2_BaseClass/DUT/Response/I_T_ResponseResult
INTERFACE I_T_ResponseResult EXTENDS KOSTAL_AF2024_Core_System.I_Interface

METHOD PUBLIC CopyTo
VAR_INPUT
	Target	: I_T_ResponseResult_CopyFrom;
END_VAR
END_METHOD

PROPERTY PUBLIC errorMessage : KOSTAL_AF2024_Core_Settings.T_MaxString_UTF8
GET
END_GET
END_PROPERTY

PROPERTY PUBLIC internalDuration : TIME
GET
END_GET
END_PROPERTY

PROPERTY PUBLIC isErrorOccured : BOOL
GET
END_GET
END_PROPERTY

PROPERTY PUBLIC isResultGood : BOOL
GET
END_GET
END_PROPERTY

END_INTERFACE

// 2_BaseClass/DUT/Response/I_T_ResponseResult_CopyFrom
INTERFACE I_T_ResponseResult_CopyFrom EXTENDS KOSTAL_AF2024_Core_System.I_Interface

METHOD PUBLIC CopyFrom
VAR_INPUT
	IN	: KOSTAL_AF2024_Core_System.I_Interface;
END_VAR
END_METHOD

END_INTERFACE

// 2_BaseClass/DUT/Response/I_T_ResponseResult_Owner
INTERFACE I_T_ResponseResult_Owner EXTENDS KOSTAL_AF2024_Core_System.I_Interface

METHOD PUBLIC clear
VAR_INPUT
END_VAR
END_METHOD

METHOD PUBLIC CopyFrom
VAR_INPUT
	IN	: KOSTAL_AF2024_Core_System.I_Interface;
END_VAR
END_METHOD

METHOD PUBLIC CopyTo
VAR_INPUT
	Target	: I_T_ResponseResult_CopyFrom;
END_VAR
END_METHOD

PROPERTY PUBLIC errorMessage :KOSTAL_AF2024_Core_Settings.T_MaxString_UTF8
GET
END_GET
SET
END_SET
END_PROPERTY

PROPERTY PUBLIC internalDuration : TIME
GET
END_GET
SET
END_SET
END_PROPERTY

PROPERTY PUBLIC isErrorOccured : BOOL
GET
END_GET
SET
END_SET
END_PROPERTY

PROPERTY PUBLIC isResultGood : BOOL
GET
END_GET
SET
END_SET
END_PROPERTY

END_INTERFACE

// 2_BaseClass/DUT/Response/T_ResponseResult
FUNCTION_BLOCK PUBLIC T_ResponseResult IMPLEMENTS I_T_ResponseResult_Owner, I_T_ResponseResult, I_T_ResponseResult_CopyFrom

VAR
	_isErrorOccured		: BOOL;
	_isResultGood			: BOOL;
	_errorMessage			: KOSTAL_AF2024_Core_Settings.T_MaxString_UTF8;
	_internalDuration	: TIME;
END_VAR

METHOD PUBLIC clear
VAR_INPUT
END_VAR


_isErrorOccured		:= FALSE;
_isResultGood			:= FALSE;
_errorMessage			:= '';
_internalDuration	:= T#0MS;
END_METHOD

METHOD PUBLIC CopyFrom
VAR_INPUT
	IN	: KOSTAL_AF2024_Core_System.I_Interface;
END_VAR

VAR
	_IN	: I_T_ResponseResult;
END_VAR

IF IN = 0 THEN RETURN;	END_IF
IF NOT __QUERYINTERFACE(IN, _IN) OR_ELSE _IN = 0 THEN RETURN;	END_IF

_isErrorOccured		:= _IN.isErrorOccured;
_isResultGood			:= _IN.isResultGood;
_errorMessage			:= _IN.errorMessage;
_internalDuration	:= _IN.internalDuration;
END_METHOD

METHOD PUBLIC CopyTo
VAR_INPUT
	Target	: I_T_ResponseResult_CopyFrom;
END_VAR

IF Target = 0 THEN RETURN;	END_IF

Target.CopyFrom(THIS^);
END_METHOD

PROPERTY PUBLIC errorMessage :KOSTAL_AF2024_Core_Settings.T_MaxString_UTF8
GET

errorMessage:= _errorMessage;
END_GET
SET

_errorMessage:= errorMessage;
END_SET
END_PROPERTY

PROPERTY PUBLIC internalDuration : TIME
GET

internalDuration:= _internalDuration;
END_GET
SET

_internalDuration:= internalDuration;
END_SET
END_PROPERTY

PROPERTY PUBLIC isErrorOccured : BOOL
GET

isErrorOccured:=	_isErrorOccured;
END_GET
SET

_isErrorOccured:=	isErrorOccured;
END_SET
END_PROPERTY

PROPERTY PUBLIC isResultGood : BOOL
GET


isResultGood:= _isResultGood;
END_GET
SET

_isResultGood:= isResultGood;
END_SET
END_PROPERTY

END_FUNCTION_BLOCK

// 2_BaseClass/POE/FB_LC
(*
|MUST EXEND
|
|TLS Parameter Initialisierung:
|================================

|https://infosys.beckhoff.de/index.php?content=../content/1031/tc3_plc_intro/index.html&id=3377440220049396176
|
|ParameterList
|The parameter list of the Tc3_IotBase library can be used to modify the size of different parameters. This modification is not possible during runtime and can only be done before compiling the code. For a better overview, only the parameter that are important for HTTP are listed in this documentation.

|Syntax
|Definition:

|VAR_GLOBAL CONSTANT Parameter_List
|    cSizeOfHttpContentType      : UDINT(32..10000);
|    cSizeOfHttpClientHostName   : UDINT(32..10000);
|    cSizeOfHttpTlsFilePaths     : UDINT(32..10000);
|    cSizeOfHttpTlsKeyFile       : UDINT(32..10000);
|    cSizeOfHttpTlsKeyPwd        : UDINT(32..10000);
|    cSizeOfHttpTlsCiphers       : UDINT(32..10000);
|    cSizeOfHttpTlsPskIdentity   : UDINT(32..10000);
|    cSizeOfHttpTlsPskKey        : UDINT(32..10000);
|END_VAR

|--------------------------|-----------------|--------------------------------------------------------------------|
|Parameter Name            |Type             |Description                                                         |
|==========================+=================+====================================================================|
|cSizeOfHttpContentType    |UDINT(32..10000) |String size definition of HTTP content type (in bytes).             |
|--------------------|-----|-----------------|--------------------------------------------------------------------|
|cSizeOfHttpClientHostName |UDINT(32..10000) |String size definition of HTTP client hostname (in bytes).          |
|--------------------|-----|-----------------|--------------------------------------------------------------------|
|cSizeOfHttpTlsFilePaths   |UDINT(32..10000) |String size definition of HTTP TLS file path (in bytes).            |
|--------------------|-----|-----------------|--------------------------------------------------------------------|
|cSizeOfHttpTlsKeyFile     |UDINT(32..10000) |String size definition of HTTP TLS key file (in bytes).             |
|--------------------|-----|-----------------|--------------------------------------------------------------------|
|cSizeOfHttpTlsKeyPwd      |UDINT(32..10000) |String size definition of HTTP TLS private key password (in bytes). |
|--------------------|-----|-----------------|--------------------------------------------------------------------|
|cSizeOfHttpTlsCiphers     |UDINT(32..10000) |String size definition of HTTP TLS cipher suites (in bytes).        |
|--------------------|-----|-----------------|--------------------------------------------------------------------|
|cSizeOfHttpTlsPskIdentity |UDINT(32..10000) |String size definition of HTTP TLS PSK identity (in bytes).         |
|--------------------|-----|-----------------|--------------------------------------------------------------------|
|cSizeOfHttpTlsPskKey      |UDINT(32..10000) |String size definition of HTTP TLS PSK (in bytes).                  |
|--------------------|-----|-----------------|--------------------------------------------------------------------|

*)
FUNCTION_BLOCK ABSTRACT FB_LC

VAR
	//Multitask Usage
	MT_Usage	: BOOL:= FALSE;;

	{region 'Client Configuration'}

		//Client Configuration request
		_HostName		: KOSTAL_AF2024_Core_Settings.T_MaxString_UTF8:= '127.0.0.1';
		_HostPort		: UINT:= 443;
		_KeepAlive	: BOOL:= FALSE;
		_TimeOut		: TIME:= T#10S;

		_TLS					: Tc3_IotBase.ST_IotSocketTls;
		_chipherSuite	: KOSTAL_AF2024_Core_Settings.T_MaxString_UTF8:= KOSTAL_AF2024_Connectivity_TLS_CipherSuite_OpenSSL.TLS_V1_2.AES128_SHA256;
		_useTLS				: BOOL:= TRUE;
		
		//Client Configuration set Variables monitored
		_HostNameSet	: KOSTAL_AF2024_Core_Settings.T_MaxString_UTF8:= '127.0.0.1';
		_HostPortSet	: UINT:= 443;

	{endregion}

	_ClientName			: KOSTAL_AF2024_Core_Settings.T_MaxString_UTF8;
	_ClientProcess	: KOSTAL_AF2024_Core_Settings.T_MaxString_UTF8;

	
	//Error without json content
	_sError_GET				: KOSTAL_AF2024_Core_Settings.T_MaxString_UTF8;
	_jsonDocError_GET	: BOOL;

	_sError_SET				: KOSTAL_AF2024_Core_Settings.T_MaxString_UTF8;
	_jsonDocError_SET	: BOOL;
	
	//
	_step		: KOSTAL_AF2024_Core_Process.FB_processStep;
	_state	: KOSTAL_AF2024_Core_Process.T_plcState;
	
	_isInit	: BOOL;
	
	_concat	: KOSTAL_AF2024_Core_StringTools.FB_Concat_UTF8;
	
	//
	_client									: Tc3_IotBase.FB_IotHttpClient;
	_clientRedirect					: BOOL:= FALSE;
	_clientCfgStep					: KOSTAL_AF2024_Core_Process.FB_processStep;
	//_clientIsDisconnecting	: BOOL;
	_clientRelease					: BOOL;
	//
	_IotHttpRequest	: Tc3_IotBase.FB_IotHttpRequest;
	_JsonParser			: Tc3_JsonXml.FB_JsonDomParser;
   _jsonDoc    		: Tc3_IotBase.SJsonValue;
	
	//
	_sUrl_Base	: KOSTAL_AF2024_Core_Settings.T_MaxString_UTF8:= URL.URI_BASE;
	_sUrl				: KOSTAL_AF2024_Core_Settings.T_MaxString_UTF8;

	//
	_ResponseResult	: T_ResponseResult;
	_sResp					: KOSTAL_AF2024_Core_Settings.T_MaxString_UTF8;

	//
	_THIS_CALLED			: E_PROCESS;
	_THIS_IN_PROCESS	: E_PROCESS;

	_ITime	: KOSTAL_AF2024_Core_GetSystemTime.I_TimeSource;

	//save to file 
	_saveFileName	: KOSTAL_AF2024_Core_Settings.T_MaxString_UTF8:= '';	//save location
	_saved				: BOOL;
	_SAVE					: BOOL;

	//Verbose
	_Verbose												: E_Verbose;

	//
	_Path_Logger									: KOSTAL_AF2024_Core_Settings.T_MaxString_UTF8;
	_File_Logger									: KOSTAL_AF2024_Core_Settings.T_MaxString_UTF8;
	_fullQualifiedFileName_Logger	: KOSTAL_AF2024_Core_Settings.T_MaxString_UTF8;
	_logger												: KOSTAL_AF2024_Core_FileLogger.FB_FileLogger;
	
	_repeatsOnFail	: UINT;
	_RepeatCount	: UINT;
	
	_AddressREPEAT: INT;
	
	_StartMessageLogged	: BOOL;
END_VAR

VAR CONSTANT
	_ADDRESS_READY	: INT:= 0;
END_VAR

METHOD PROTECTED _getResponseResultFromJson : KOSTAL_AF2024_Core_Settings.T_MaxString_UTF8

VAR_INPUT
	IN	: Tc3_IotBase.SJsonValue;
	OUT	: REFERENCE TO T_ResponseResult;
END_VAR

VAR
	_isErrorOccured: BOOL;
	_isResultGood: BOOL;
	_errorMessage	: KOSTAL_AF2024_Core_Settings.T_MaxString_UTF8;
	_internalDuration	: TIME;
	
	_resp	: KOSTAL_AF2024_Core_Settings.T_MaxString_UTF8;
END_VAR
	
IF IN = 0 THEN _getResponseResultFromJson:= ';_getResponseBodyFromJson - IN Parameter is empty';	RETURN;	END_IF
IF NOT __ISVALIDREF(OUT) THEN _getResponseResultFromJson:= '_getResponseBodyFromJson - OUT Parameter is invalid';	RETURN;	END_IF

_getResponseResultFromJson:= '';
OUT.clear();

_resp:= _PARSE_BOOL(IN, RESPONSE_BODY.isErrorOccured, _isErrorOccured);
IF _resp = '' 											THEN	OUT.isErrorOccured:= _isErrorOccured;	
ELSIF _getResponseResultFromJson = ''	THEN _getResponseResultFromJson:= _resp;
END_IF

_resp:= _PARSE_BOOL(IN, RESPONSE_BODY.isResultGood, _isResultGood);
IF _resp = '' 											THEN	OUT.isResultGood:= _isResultGood;
ELSIF _getResponseResultFromJson = ''	THEN _getResponseResultFromJson:= _resp;
END_IF

_resp:= _PARSE_STRING(IN, RESPONSE_BODY.errorMessage, _errorMessage);
IF _resp = '' THEN	OUT.errorMessage:= _errorMessage;
ELSIF _getResponseResultFromJson = ''	THEN _getResponseResultFromJson:= _resp;
END_IF

_resp:= _PARSE_TIME(IN, RESPONSE_BODY.internalDuration, _internalDuration);
IF _resp = '' THEN	OUT.internalDuration:= _internalDuration;
ELSIF _getResponseResultFromJson = ''	THEN _getResponseResultFromJson:= _resp;
END_IF
END_METHOD

(*
| return a Json Value with access to an Array
*)
METHOD PROTECTED _PARSE_ARRAY : KOSTAL_AF2024_Core_Settings.T_MaxString_UTF8

VAR_INPUT
	IN			: Tc3_IotBase.SJsonValue;
	Member	: KOSTAL_AF2024_Core_Settings.T_MaxString_UTF8;	
	Q				: REFERENCE TO Tc3_IotBase.SJsonValue;	
	
END_VAR

VAR
	_J	:	Tc3_IotBase.SJsonValue;
END_VAR


IF IN = 0 THEN _PARSE_ARRAY:= Tc2_Standard.CONCAT(Member,  ';_PARSE_ARRAY - IN Parameter is empty');	RETURN;	END_IF
IF NOT __ISVALIDREF(Q) THEN _PARSE_ARRAY:= Tc2_Standard.CONCAT(Member,  ';_PARSE_ARRAY - Q Parameter is invalid');	RETURN;	END_IF


_PARSE_ARRAY:= '';
_J:= 0;


IF NOT _JsonParser.HasMember(IN, Member) THEN	Q:= 0; _PARSE_ARRAY:= Tc2_Standard.CONCAT(Member,  ';_PARSE_ARRAY - no member');	RETURN;	END_IF

_J:= _JsonParser.FindMember(IN,	Member);

IF _J = 0 THEN	Q:= 0;	_PARSE_ARRAY:=  Tc2_Standard.CONCAT(Member,  ';_PARSE_ARRAY - no member');	RETURN;	END_IF

IF NOT _JsonParser.IsArray(_J) THEN Q:= 0;	_PARSE_ARRAY:=  Tc2_Standard.CONCAT(Member,  ';_PARSE_ARRAY - is not an Array');	RETURN;	END_IF

Q:= _J;	

IF _JsonParser.IsNull(_J) THEN	Q:= 0; _PARSE_ARRAY:= Tc2_Standard.CONCAT(Member,  ';_PARSE_ARRAY - no content'); RETURN;	END_IF
END_METHOD

METHOD PROTECTED _PARSE_BOOL : KOSTAL_AF2024_Core_Settings.T_MaxString_UTF8

VAR_INPUT
	IN			: Tc3_IotBase.SJsonValue;
	Member	: KOSTAL_AF2024_Core_Settings.T_MaxString_UTF8;	
	Q				: REFERENCE TO BOOL;
END_VAR

VAR
	_J	:	Tc3_IotBase.SJsonValue;
END_VAR

IF IN = 0 THEN _PARSE_BOOL:= Tc2_Standard.CONCAT(Member,  ';_PARSE_BOOL - IN Parameter is empty');	RETURN;	END_IF
IF NOT __ISVALIDREF(Q) THEN _PARSE_BOOL:= Tc2_Standard.CONCAT(Member,  ';_PARSE_BOOL - Q Parameter is invalid');	RETURN;	END_IF


_PARSE_BOOL:= '';


IF NOT _JsonParser.HasMember(IN, Member) THEN	Q:= FALSE; _PARSE_BOOL:= Tc2_Standard.CONCAT(Member,  ';_PARSE_BOOL - no member');	RETURN;	END_IF

_J:= _JsonParser.FindMember(IN,	Member);

IF _J = 0 THEN	_PARSE_BOOL:=  Tc2_Standard.CONCAT(Member,  ';_PARSE_BOOL - no member');	RETURN;	END_IF

IF 		_JsonParser.IsNull(_J) 		THEN	Q:= FALSE; 
ELSIF _JsonParser.IsBool(_J) 		THEN	Q:= _JsonParser.GetBool(v:= _J);	
ELSIF _JsonParser.IsNumber(_J)	THEN	Q:=  UDINT_TO_BOOL(_JsonParser.GetUint(_J));
ELSE																	Q:= FALSE; _PARSE_BOOL:= Tc2_Standard.CONCAT(Member,  ';_PARSE_BOOL - not BOOL');
END_IF
END_METHOD

METHOD PROTECTED _PARSE_BYTE : KOSTAL_AF2024_Core_Settings.T_MaxString_UTF8

VAR_INPUT
	IN			: Tc3_IotBase.SJsonValue;
	Member	: KOSTAL_AF2024_Core_Settings.T_MaxString_UTF8;	
	Q				: REFERENCE TO BYTE;
END_VAR

VAR
	_J	:	Tc3_IotBase.SJsonValue;
END_VAR

IF IN = 0 THEN _PARSE_BYTE:= Tc2_Standard.CONCAT(Member,  ';_PARSE_BYTE - IN Parameter is empty');	RETURN;	END_IF
IF NOT __ISVALIDREF(Q) THEN _PARSE_BYTE:= Tc2_Standard.CONCAT(Member,  ';_PARSE_BYTE - Q Parameter is invalid');	RETURN;	END_IF


_PARSE_BYTE:= '';

IF NOT _JsonParser.HasMember(IN, Member) THEN	Q:= 0; _PARSE_BYTE:= Tc2_Standard.CONCAT(Member,  ';_PARSE_BYTE - no member');	RETURN;	END_IF

_J:= _JsonParser.FindMember(IN,	Member);

IF _J = 0 THEN	Q:= 0; _PARSE_BYTE:=  Tc2_Standard.CONCAT(Member,  ';_PARSE_BYTE - no member');	RETURN;	END_IF

IF _JsonParser.IsNull(_J) THEN	Q:= 0; RETURN;	END_IF

IF NOT _JsonParser.IsNumber(_J) THEN	Q:= 0; _PARSE_BYTE:= Tc2_Standard.CONCAT(Member,  ';_PARSE_BYTE - not BYTE/Number');	RETURN;	END_IF

Q	:= UDINT_TO_BYTE(_JsonParser.GetUint(v:= _J));
END_METHOD

METHOD PROTECTED _PARSE_DINT : KOSTAL_AF2024_Core_Settings.T_MaxString_UTF8

VAR_INPUT
	IN			: Tc3_IotBase.SJsonValue;
	Member	: KOSTAL_AF2024_Core_Settings.T_MaxString_UTF8;	
	Q				: REFERENCE TO DINT;
END_VAR

VAR
	_J	:	Tc3_IotBase.SJsonValue;
END_VAR

IF IN = 0 THEN _PARSE_DINT:= Tc2_Standard.CONCAT(Member,  ';_PARSE_DINT - IN Parameter is empty');	RETURN;	END_IF
IF NOT __ISVALIDREF(Q) THEN _PARSE_DINT:= Tc2_Standard.CONCAT(Member,  ';_PARSE_DINT - Q Parameter is invalid');	RETURN;	END_IF


_PARSE_DINT:= '';

IF NOT _JsonParser.HasMember(IN, Member) THEN	Q:= 0; _PARSE_DINT:= Tc2_Standard.CONCAT(Member,  ';_PARSE_DINT - no member');	RETURN;	END_IF

_J:= _JsonParser.FindMember(IN,	Member);

IF _J = 0 THEN	Q:= 0; _PARSE_DINT:=  Tc2_Standard.CONCAT(Member,  ';_PARSE_DINT - no member');	RETURN;	END_IF

IF _JsonParser.IsNull(_J) THEN	Q:= 0; RETURN;	END_IF

IF NOT _JsonParser.IsNumber(_J) THEN	Q:= 0; _PARSE_DINT:= Tc2_Standard.CONCAT(Member,  ';_PARSE_DINT - not DINT/Number');	RETURN;	END_IF

Q	:= _JsonParser.GetInt(v:= _J);
END_METHOD

(*
| return a Json Value with access to an Array
*)
METHOD PROTECTED _PARSE_JSON : KOSTAL_AF2024_Core_Settings.T_MaxString_UTF8

VAR_INPUT
	IN			: Tc3_IotBase.SJsonValue;
	Member	: KOSTAL_AF2024_Core_Settings.T_MaxString_UTF8;	
	Q				: REFERENCE TO Tc3_IotBase.SJsonValue;	
	
END_VAR

VAR
	_J	:	Tc3_IotBase.SJsonValue;
END_VAR


IF IN = 0 THEN _PARSE_JSON:= Tc2_Standard.CONCAT(Member,  ';_PARSE_JSON - IN Parameter is empty');	RETURN;	END_IF
IF NOT __ISVALIDREF(Q) THEN _PARSE_JSON:= Tc2_Standard.CONCAT(Member,  ';_PARSE_JSON - Q Parameter is invalid');	RETURN;	END_IF


_PARSE_JSON:= '';
_J:= 0;


IF NOT _JsonParser.HasMember(IN, Member) THEN	Q:= 0; _PARSE_JSON:= Tc2_Standard.CONCAT(Member,  ';_PARSE_JSON - no member');	RETURN;	END_IF

_J:= _JsonParser.FindMember(IN,	Member);

IF _J = 0 THEN	Q:= 0;	_PARSE_JSON:=  Tc2_Standard.CONCAT(Member,  ';_PARSE_JSON - no member');	RETURN;	END_IF

Q:= _J;	

IF _JsonParser.IsNull(_J) THEN	Q:= 0; _PARSE_JSON:= Tc2_Standard.CONCAT(Member,  ';_PARSE_JSON - no content'); RETURN;	END_IF
END_METHOD

METHOD PROTECTED _PARSE_STRING : KOSTAL_AF2024_Core_Settings.T_MaxString_UTF8

VAR_INPUT
	IN			: Tc3_IotBase.SJsonValue;
	Member	: KOSTAL_AF2024_Core_Settings.T_MaxString_UTF8;	
	Q				: REFERENCE TO KOSTAL_AF2024_Core_Settings.T_MaxString_UTF8;
END_VAR

VAR
	_J	:	Tc3_IotBase.SJsonValue;
END_VAR

IF IN = 0 THEN _PARSE_STRING:= Tc2_Standard.CONCAT(Member,  ';_PARSE_STRING - IN Parameter is empty');	RETURN;	END_IF
IF NOT __ISVALIDREF(Q) THEN _PARSE_STRING:= Tc2_Standard.CONCAT(Member,  ';_PARSE_STRING - Q Parameter is invalid');	RETURN;	END_IF


_PARSE_STRING:= '';


IF NOT _JsonParser.HasMember(IN, Member) THEN	Q:= ''; _PARSE_STRING:= Tc2_Standard.CONCAT(Member,  ';_PARSE_STRING - no member');	RETURN;	END_IF

_J:= _JsonParser.FindMember(IN,	Member);

IF _J = 0 THEN	Q:= ''; _PARSE_STRING:=  Tc2_Standard.CONCAT(Member,  ';_PARSE_STRING - no member');	RETURN;	END_IF

IF _JsonParser.IsNull(_J) THEN	Q:= ''; RETURN;	END_IF

IF NOT _JsonParser.IsString(_J) THEN	Q:= ''; _PARSE_STRING:= Tc2_Standard.CONCAT(Member,  ';_PARSE_STRING - not STRING');	RETURN;	END_IF

Q:= _JsonParser.GetString(v:= _J);
END_METHOD

METHOD PROTECTED _PARSE_TIME : KOSTAL_AF2024_Core_Settings.T_MaxString_UTF8

VAR_INPUT
	IN			: Tc3_IotBase.SJsonValue;
	Member	: KOSTAL_AF2024_Core_Settings.T_MaxString_UTF8;	
	Q				: REFERENCE TO TIME;
END_VAR

VAR
	_J	:	Tc3_IotBase.SJsonValue;
	_num: ULINT;
END_VAR

IF IN = 0 THEN _PARSE_TIME:= Tc2_Standard.CONCAT(Member,  ';_PARSE_TIME - IN Parameter is empty');	RETURN;	END_IF
IF NOT __ISVALIDREF(Q) THEN _PARSE_TIME:= Tc2_Standard.CONCAT(Member,  ';_PARSE_TIME - Q Parameter is invalid');	RETURN;	END_IF


_PARSE_TIME:= '';

IF NOT _JsonParser.HasMember(IN, Member) THEN	Q:= T#0MS; _PARSE_TIME:= Tc2_Standard.CONCAT(Member,  ';_PARSE_TIME - no member');	RETURN;	END_IF

_J:= _JsonParser.FindMember(IN,	Member);

IF _J = 0 THEN	Q:= T#0MS; _PARSE_TIME:=  Tc2_Standard.CONCAT(Member,  ';_PARSE_TIME - no member');	RETURN;	END_IF

IF _JsonParser.IsNull(_J) THEN	Q:= T#0MS; RETURN;	END_IF

IF NOT _JsonParser.IsNumber(_J) THEN	Q:= T#0MS; _PARSE_TIME:= Tc2_Standard.CONCAT(Member,  ';_PARSE_TIME - not TIME');	RETURN;	END_IF

_num	:= _JsonParser.GetUint64(v:= _J);

Q := ULINT_TO_TIME(_num);
END_METHOD

METHOD PROTECTED _PARSE_UDINT : KOSTAL_AF2024_Core_Settings.T_MaxString_UTF8

VAR_INPUT
	IN			: Tc3_IotBase.SJsonValue;
	Member	: KOSTAL_AF2024_Core_Settings.T_MaxString_UTF8;	
	Q				: REFERENCE TO UDINT;
END_VAR

VAR
	_J	:	Tc3_IotBase.SJsonValue;
END_VAR

IF IN = 0 THEN _PARSE_UDINT:= Tc2_Standard.CONCAT(Member,  ';_PARSE_UDINT - IN Parameter is empty');	RETURN;	END_IF
IF NOT __ISVALIDREF(Q) THEN _PARSE_UDINT:= Tc2_Standard.CONCAT(Member,  ';_PARSE_UDINT - Q Parameter is invalid');	RETURN;	END_IF


_PARSE_UDINT:= '';

IF NOT _JsonParser.HasMember(IN, Member) THEN	Q:= 0; _PARSE_UDINT:= Tc2_Standard.CONCAT(Member,  ';_PARSE_UDINT - no member');	RETURN;	END_IF

_J:= _JsonParser.FindMember(IN,	Member);

IF _J = 0 THEN	Q:= 0; _PARSE_UDINT:=  Tc2_Standard.CONCAT(Member,  ';_PARSE_UDINT - no member');	RETURN;	END_IF

IF _JsonParser.IsNull(_J) THEN	Q:= 0; RETURN;	END_IF

IF NOT _JsonParser.IsNumber(_J) THEN	Q:= 0; _PARSE_UDINT:= Tc2_Standard.CONCAT(Member,  ';_PARSE_UDINT - not UDINT/Number');	RETURN;	END_IF

Q	:= _JsonParser.GetUint(v:= _J);
END_METHOD

METHOD PROTECTED _PARSE_ULINT : KOSTAL_AF2024_Core_Settings.T_MaxString_UTF8

VAR_INPUT
	IN			: Tc3_IotBase.SJsonValue;
	Member	: KOSTAL_AF2024_Core_Settings.T_MaxString_UTF8;	
	Q				: REFERENCE TO ULINT;
END_VAR

VAR
	_J	:	Tc3_IotBase.SJsonValue;
END_VAR

IF IN = 0 THEN _PARSE_ULINT:= Tc2_Standard.CONCAT(Member,  ';_PARSE_ULINT - IN Parameter is empty');	RETURN;	END_IF
IF NOT __ISVALIDREF(Q) THEN _PARSE_ULINT:= Tc2_Standard.CONCAT(Member,  ';_PARSE_ULINT - Q Parameter is invalid');	RETURN;	END_IF


_PARSE_ULINT:= '';

IF NOT _JsonParser.HasMember(IN, Member) THEN	Q:= 0; _PARSE_ULINT:= Tc2_Standard.CONCAT(Member,  ';_PARSE_ULINT - no member');	RETURN;	END_IF

_J:= _JsonParser.FindMember(IN,	Member);

IF _J = 0 THEN	Q:= 0; _PARSE_ULINT:=  Tc2_Standard.CONCAT(Member,  ';_PARSE_ULINT - no member');	RETURN;	END_IF

IF _JsonParser.IsNull(_J) THEN	Q:= 0; RETURN;	END_IF

IF NOT _JsonParser.IsNumber(_J) THEN	Q:= 0; _PARSE_ULINT:= Tc2_Standard.CONCAT(Member,  ';_PARSE_ULINT - _PARSE_ULINT - not ULINT/Number');	RETURN;	END_IF

Q	:= _JsonParser.GetUint64(v:= _J);
END_METHOD

METHOD PROTECTED _00_clientCfg 

VAR
	_c	: KOSTAL_AF2024_Core_StringTools.FB_Concat;
END_VAR

IF _step.toggle THEN
	_clientCfgStep.init();
END_IF


_clientCfgStep.Header();

CASE _clientCfgStep.actual OF

	0:	IF		_CfgHasChanged()				THEN	_clientRelease:= FALSE;	_clientCfgStep.INC();
			ELSIF	_client.bError					THEN	_clientRelease:= FALSE;	_clientCfgStep.INC();
			ELSIF	NOT _client.bConfigured	THEN	_clientRelease:= FALSE;	_clientCfgStep.INC();
			ELSIF	NOT _clientRelease			THEN	_clientCfgStep.INC();
			ELSE 													_step.INC();
			END_IF

	
	1:	_client.Disconnect();
			
			
			_state.clear();
			_state.busy:= TRUE;
			_state.description:= "Reconfiguration runs ...";
			
			IF NOT _client.bConfigured THEN	
				_CfgChange();	
				_clientCfgStep.INC();	
			END_IF
			
	2:	
			_state.clear();
			_state.busy:= TRUE;
			_state.description:= "wait for Reconfiguration completed ...";
		
			_client.Execute();
			
			IF _client.bConfigured THEN	
				_clientRelease:= TRUE;
				_step.INC();
			END_IF

			
ELSE
		
	_state.clear();
	
	_state.fail:= TRUE;
	
	_c.clear();
	_c.addContent("_clientCfgStep ");
	_c.addContent(INT_TO_WSTRING(_clientCfgStep.actual));
	_c.addContent(" do not exist...");
	
	_state.description:= _c.getResult();
	_c.clear();
	
	_state.finish:= TRUE;


END_CASE
END_METHOD

METHOD PROTECTED _01_Ready : BOOL
VAR_INPUT
END_VAR

IF _step.toggle THEN
	
	//_client.Disconnect();
	_THIS_IN_PROCESS:=  E_PROCESS.idle;

END_IF

_01_Ready:= TRUE;//_client.bConfigured;

IF NOT _01_Ready THEN
	_state.clear();
	_state.fail:= TRUE;
	_state.description:= "Client not configured";
END_IF

(*
IF _ClientName = '' THEN

	_state.clear();
	_state.fail:= TRUE;
	_state.description:= 'No Client Name defined - like SPSPCxxx';
	
ELSIF _ClientProcess = '' THEN

	_state.clear();
	_state.fail:= TRUE;
	_state.description:= 'No Client Process defined - like ASSxx';

ELSE

	_01_Ready:= TRUE;

END_IF
*)
END_METHOD

METHOD PROTECTED _10_finishFail
VAR_INPUT
END_VAR



IF _step.toggle THEN
	_JsonParser.NewDocument();
END_IF

_state.finish:= TRUE;
_state.pass:= FALSE;
_state.fail:= TRUE;
END_METHOD

METHOD PROTECTED _10_finishPass
VAR_INPUT
END_VAR



IF _step.toggle THEN
	_JsonParser.NewDocument();
END_IF

_state.clear();
_state.finish:= TRUE;
_state.pass:= TRUE;
END_METHOD

METHOD PROTECTED _10_GET
VAR_INPUT
END_VAR

IF _step.toggle THEN
	_AddressREPEAT:= _step.actual;
END_IF


IF _IotHttpRequest.SendRequest
	(
		sUri:= _sUrl,
		fbClient:= _Client,
		eRequestType:= Tc3_IotBase.ETcIotHttpRequestType.HTTP_GET,
		pContent:= 0,
		nContentSize:= 0,
		fbHeader:= 0
	) THEN	

	_state.description:= ""; 

	_step.INC();	

ELSE
	
	_state.description:= "wait for IotHttpRequest.SendRequest";

END_IF
END_METHOD

METHOD PROTECTED _10_GET_CTRL
VAR_INPUT
END_VAR
IF _step.toggle THEN
	;
END_IF

IF _IotHttpRequest.bBusy THEN

	_state.description:= "_IotHttpRequest is busy... wait for finish;"; 

ELSIF _IotHttpRequest.bError THEN

	_state.clear();
	_state.finish:= TRUE;
	_state.fail:= TRUE;
	_state.description:= Tc2_Standard.WCONCAT("_IotHttpRequest returns an error Number:;", DINT_TO_WSTRING(_IotHttpRequest.eErrorId)); 

	IF (_RepeatCount < _repeatsOnFail) THEN	
		_RepeatCount:= _RepeatCount + 1;
		_step.set(_AddressREPEAT);
	END_IF

(*ELSIF _IotHttpRequest.nStatusCode < 200 OR _IotHttpRequest.nStatusCode > 299 THEN


	_RepeatCount:= 0;

	_state.clear();
	_state.setUnique_finish();
	_state.fail:= TRUE;
	_state.description:= Tc2_Standard.CONCAT('_IotHttpRequest returns a status Number:;', UINT_TO_STRING(_IotHttpRequest.nStatusCode)); 
*)

ELSIF _IotHttpRequest.nContentSize = 0 THEN

	_RepeatCount:= 0;

	_state.clear();
	_state.finish:= TRUE;
	_state.fail:= TRUE;
	_state.description:= "_IotHttpRequest returns no content"; 

ELSE

		_RepeatCount:= 0;
		

		_jsonDoc:= _IotHttpRequest.GetJsonDomContent(_JsonParser);

		IF _jsonDoc = 0 THEN

			_IotHttpRequest.GetContent(ADR(_sError_GET), SIZEOF(_sError_GET), TRUE);

			IF _logger.enabled AND NOT _jsonDocError_GET THEN 

				_logger.addLine(TO_WSTRING(_sError_GET));	
				_jsonDocError_GET:= TRUE;	

			END_IF

		ELSE

			_jsonDocError_GET:= FALSE;

		END_IF
		
		
	_step.INC();

END_IF
END_METHOD

METHOD PROTECTED _10_GET_ResponseResult
VAR_INPUT
	logUri	: BOOL;
END_VAR

IF _step.toggle THEN
		_VerboseHandler(_JsonParser.GetDocumentLength() <> 0, 'GET', logUri);
END_IF


IF _SAVE THEN

	_state.description:= Tc2_Standard.WCONCAT("Wait for saved the Json Document to : ", TO_WSTRING(_saveFileName));
 
ELSIF _jsonDoc = 0 THEN

	_state.clear();
	_state.finish:= TRUE;
	_state.fail:= TRUE;
	_state.description:= "no Json response available";
	
ELSE
	
	_sResp:= _getResponseResultFromJson(_jsonDoc,_ResponseResult);
	

	_step.INC();

END_IF
END_METHOD

METHOD PROTECTED _10_GET_ResponseResult_CTRL
VAR_INPUT
END_VAR

IF _step.toggle THEN
	;
END_IF


IF _sResp <> '' THEN

	_state.clear();
	_state.finish:= TRUE;
	_state.fail:= TRUE;
	_state.description:= Tc2_Standard.WCONCAT("Response is incomplete;", TO_WSTRING(_sResp));
	
ELSIF _ResponseResult.isErrorOccured THEN
	
	_state.clear();
	_state.finish:= TRUE;
	_state.fail:= TRUE;
	_state.description:= Tc2_Standard.WCONCAT("Response failed;", TO_WSTRING(_ResponseResult.errorMessage));

ELSE
	

	_step.INC();

END_IF
END_METHOD

METHOD PROTECTED _10_SET
VAR_INPUT
	logUri	: BOOL;
END_VAR
				
IF _step.toggle THEN
	_AddressREPEAT:= _step.actual;
	_VerboseHandler(_JsonParser.GetDocumentLength() <> 0, 'SET', logUri);
END_IF


IF _SAVE THEN

	_state.description:= Tc2_Standard.WCONCAT("Wait for saved the Json Document to : ", TO_WSTRING(_saveFileName));
 
ELSIF _IotHttpRequest.SendJsonDomRequest
	(
		sUri:= _sUrl,
		fbClient:= _Client,
		fbJson:= _JsonParser,
		eRequestType:= Tc3_IotBase.ETcIotHttpRequestType.HTTP_POST,
		fbHeader:= 0
	) THEN	

	_state.description:= ""; 

	_step.INC();	

ELSE
	
	_state.description:= "wait for IotHttpRequest.SendJsonDomRequest";

END_IF
END_METHOD

METHOD PROTECTED _10_SET_CTRL
VAR_INPUT
END_VAR
  
IF _step.toggle THEN
	;
END_IF

IF _IotHttpRequest.bBusy THEN

	_state.description:= "_IotHttpRequest is busy... wait for finish;"; 

ELSIF _IotHttpRequest.bError THEN

	_state.clear();
	_state.finish:= TRUE;
	_state.fail:= TRUE;
	_state.description:= Tc2_Standard.WCONCAT("_IotHttpRequest returns an error Number:;", DINT_TO_WSTRING(_IotHttpRequest.eErrorId)); 

	IF (_RepeatCount < _repeatsOnFail) THEN	
		_RepeatCount:= _RepeatCount + 1;
		_step.set(_AddressREPEAT);
	END_IF

(*ELSIF _IotHttpRequest.nStatusCode < 200 OR _IotHttpRequest.nStatusCode > 299 THEN

	_RepeatCount:= 0;

	_state.clear();
	_state.setUnique_finish();
	_state.fail:= TRUE;
	_state.description:= Tc2_Standard.CONCAT('_IotHttpRequest returns a status Number:;', UINT_TO_STRING(_IotHttpRequest.nStatusCode)); 
*)

ELSE

		_RepeatCount:= 0;


		_jsonDoc:= _IotHttpRequest.GetJsonDomContent(_JsonParser);

		IF _jsonDoc = 0 THEN

			_IotHttpRequest.GetContent(ADR(_sError_SET), SIZEOF(_sError_SET), TRUE);

			IF _logger.enabled AND NOT _jsonDocError_SET THEN 

				_logger.addLine(TO_WSTRING(_sError_SET));	
				_jsonDocError_SET:= TRUE;	

			END_IF

		ELSE

			_jsonDocError_SET:= FALSE;

		END_IF
		
		
	_step.INC();

END_IF
END_METHOD

METHOD PROTECTED _99_stepError
VAR
	_c	:	KOSTAL_AF2024_Core_StringTools.FB_Concat;
END_VAR

_state.clear();

_state.fail:= TRUE;

_c.clear();
_c.addContent("step ");
_c.addContent(INT_TO_WSTRING(_step.actual));
_c.addContent(" do not exist...");

_state.description:= _c.getResult();
_c.clear();

_state.finish:= TRUE;
END_METHOD

METHOD PROTECTED _CfgChange
VAR_INPUT
END_VAR


_HostNameSet:= _HostName; 
_HostPortSet:= _HostPort;

IF _useTLS THEN	

	_TLS.bNoServerCertCheck:= TRUE;
	_TLS.sCiphers:= _chipherSuite;
	_client.stTLS	:= _TLS;	

END_IF
END_METHOD

METHOD PROTECTED _CfgHasChanged : BOOL
VAR_INPUT
END_VAR

_CfgHasChanged:= (_HostNameSet <> _HostName) 
							OR (_HostPortSet <> _HostPort);
END_METHOD

METHOD PROTECTED _deviceDefine

_client.sHostName							:= _HostNameSet;	//Client Configuration set Variables monitored
_client.nHostPort							:= _HostPortSet;	//Client Configuration set Variables monitored

_client.bKeepAlive						:= _KeepAlive;
_client.tConnectionTimeout		:= _TimeOut;

//client connecting
IF _clientRelease THEN	_client.Execute();	END_IF


_saved:= _JsonParser.SaveDocumentToFile(_saveFileName, _SAVE); 
IF _saved THEN _SAVE:= FALSE;	END_IF

IF NOT _isInit THEN
	_concat.clear();
	_concat.addContent(_Path_Logger);
	_concat.addContent(_File_Logger);
	_concat.addContent('_URL');
	_logger.Path:= _concat.getResult(); 
	_concat.clear();
END_IF

_logger.enabled:= _Verbose <> E_Verbose.none;
_logger.linkTimeSource(_ITime);
_logger.FBmain();

_logStartMessage();
END_METHOD

METHOD PROTECTED _logStartMessage

VAR
	_c	: KOSTAL_AF2024_Core_StringTools.FB_Concat;
	_stVersion: ST_LibVersion;
END_VAR

IF NOT _StartMessageLogged THEN

	IF _ITime = 0 THEN	;
	ELSIF NOT _ITime.Valid THEN	;
	ELSIF NOT _logger.enabled THEN	;
	ELSE

		_stVersion:= F_GetVersion();
		
		_c.clear();
		_c.addContent(F_GetTitle());
		_c.addContent(";");
		_c.addContent("Version:");
		_c.addContent(UINT_TO_WSTRING(_stVersion.iMajor));		
		_c.addContent(".");
		_c.addContent(UINT_TO_WSTRING(_stVersion.iMinor));		
		_c.addContent(".");
		_c.addContent(UINT_TO_WSTRING(_stVersion.iBuild));		
		_c.addContent(".");
		_c.addContent(UINT_TO_WSTRING(_stVersion.iRevision));		
		_c.addContent(";");
		_c.addContent("=START=");
		_logger.addLine(_c.getResult());
		_c.clear();
		_StartMessageLogged:= TRUE;

	END_IF

END_IF
END_METHOD

METHOD PROTECTED _UriGet : KOSTAL_AF2024_Core_Settings.T_MaxString_UTF8
VAR_INPUT
	Extension	: KOSTAL_AF2024_Core_Settings.T_MaxString_UTF8;
END_VAR

_UriGet:= Tc2_Standard.CONCAT(_sUrl_Base, Extension);
END_METHOD

(*
| Returns the Url with replaced Placeholders
*)
METHOD PROTECTED _UrlReplace

VAR_INPUT
	IN		:	REFERENCE TO KOSTAL_AF2024_Core_Settings.T_MaxString_UTF8;
	Key		: KOSTAL_AF2024_Core_Settings.T_MaxString_UTF8;
	Value	: KOSTAL_AF2024_Core_Settings.T_MaxString_UTF8;
END_VAR

VAR
	_work :	KOSTAL_AF2024_Core_Settings.T_MaxString_UTF8;
END_VAR
IF NOT __ISVALIDREF(IN) THEN RETURN;	END_IF

_work:= IN;

_work:= KOSTAL_AF2024_Core_StringTools.F_Replace_UTF8(_work, Key, Value, -1);

IN:= _work;
END_METHOD

METHOD PROTECTED _VerboseHandler : BOOL

VAR_INPUT
	withContent	: BOOL;	
	Extension		: STRING;
	logUri			: BOOL;
END_VAR

VAR
	_TS	: Tc2_Utilities.TIMESTRUCT;
	_TimeStamp	:	KOSTAL_AF2024_Core_Settings.T_MaxString_UTF8;	
END_VAR

_VerboseHandler:= FALSE;

_TS:= _ITime.GetTimeStruct();

IF _ITime <> 0 THEN	_TimeStamp:= Tc2_Utilities.SYSTEMTIME_TO_STRING(_TS);	ELSE _TimeStamp:= '';	END_IF	


_TimeStamp:= KOSTAL_AF2024_Core_StringTools.F_Replace_UTF8(_TimeStamp, ':','-', -1);

//Save Request	
IF UINT_TO_BOOL((INT_TO_WORD(_Verbose) AND 16#01)) THEN

	IF logUri THEN
//		set in _deviceDefine()		
//		_concat.clear();
//		_concat.new(3);
//		_concat.addContent(1, _Path_Logger);
//		_concat.addContent(2, _File_Logger);
//		_concat.addContent(3, '_URL');
//		_logger.fileName:= _concat.getResult(); 
	
		_logger.addLine(TO_WSTRING(_sUrl));
	END_IF
	
	IF withContent THEN
		_concat.clear();
		_concat.addContent(_Path_Logger);
		_concat.addContent(_File_Logger);
		_concat.addContent('_');
		_concat.addContent(Extension);
		_concat.addContent('_');
		_concat.addContent(_TimeStamp);
		_concat.addContent('.json');
		_fullQualifiedFileName_Logger:= _concat.getResult();
		_concat.clear();
	
		_saveFileName:= _fullQualifiedFileName_Logger;
		_SAVE:= TRUE;
	END_IF
	
	_VerboseHandler:= TRUE;

END_IF
END_METHOD

PROPERTY PUBLIC ClientName : KOSTAL_AF2024_Core_Settings.T_MaxString_UTF8
GET

ClientName:= _ClientName;
END_GET
SET

_ClientName:= ClientName;
END_SET
END_PROPERTY

PROPERTY PUBLIC ClientProcess : KOSTAL_AF2024_Core_Settings.T_MaxString_UTF8
GET

ClientProcess:= _ClientProcess;
END_GET
SET

_ClientProcess:= ClientProcess;
END_SET
END_PROPERTY

PROPERTY PUBLIC HostName : KOSTAL_AF2024_Core_Settings.T_MaxString_UTF8
GET

HostName:= _HostName;
END_GET
SET

_HostName:= HostName;
END_SET
END_PROPERTY

PROPERTY PUBLIC HostPort : UINT
GET

HostPort:= _HostPort;
END_GET
SET

_HostPort:= HostPort;
END_SET
END_PROPERTY

PROPERTY HTTP_Statuscode : UXINT
GET

HTTP_Statuscode:= _IotHttpRequest.nStatusCode;
END_GET
END_PROPERTY

(*
| Retunrs the Process which is in use
*)
PROPERTY IN_PROCESS : E_PROCESS
GET

IN_PROCESS := _THIS_IN_PROCESS;
END_GET
END_PROPERTY

(*
	Default = TRUE
*)
PROPERTY PUBLIC KeepAlive : BOOL
GET

KeepAlive:= _KeepAlive;
END_GET
SET

_KeepAlive:= KeepAlive;
END_SET
END_PROPERTY

PROPERTY PUBLIC repeatsOnFail : UINT
GET

repeatsOnFail:= _repeatsOnFail;
END_GET
SET

_repeatsOnFail:= repeatsOnFail;
END_SET
END_PROPERTY

PROPERTY State : KOSTAL_AF2024_Core_Process.I_T_plcState
GET

State := _state;
END_GET
END_PROPERTY

(*
	Default = T#10s
*)
PROPERTY PUBLIC TimeOut : TIME
GET

TimeOut:= _TimeOut;
END_GET
SET

_TimeOut:= TimeOut;
END_SET
END_PROPERTY

(*
| Interface LineCintrol Web Service Duration
*)
PROPERTY WS_Duration : TIME
GET

WS_Duration:=	_ResponseResult.internalDuration;
END_GET
END_PROPERTY

METHOD PUBLIC FBmain
VAR_INPUT
END_VAR

IF _THIS_CALLED = E_PROCESS.idle THEN
	
	_FBmain();
	
END_IF

_THIS_CALLED:= E_PROCESS.idle;
END_METHOD

METHOD PUBLIC GetTimeStamp : KOSTAL_AF2024_Core_Settings.T_MaxString_UTF8

IF _ITime <> 0 THEN GetTimeStamp:= '';	RETURN;	END_IF

_concat.clear();

_concat.addContent
	(KOSTAL_AF2024_Core_StringTools.F_FormatMask_UTF8
			(	WORD_TO_STRING(_ITime.TimeStruct.Year), 
				'2000', KOSTAL_AF2024_Core_StringTools.E_ALIGNMENT.RIGHT)); 

_concat.addContent
	('-'); 

_concat.addContent
	(KOSTAL_AF2024_Core_StringTools.F_FormatMask_UTF8
			(	WORD_TO_STRING(_ITime.TimeStruct.Month), 
				'00', KOSTAL_AF2024_Core_StringTools.E_ALIGNMENT.RIGHT)); 

_concat.addContent
	('-'); 

_concat.addContent
	(KOSTAL_AF2024_Core_StringTools.F_FormatMask_UTF8
			(	WORD_TO_STRING(_ITime.TimeStruct.Day), 
				'00', KOSTAL_AF2024_Core_StringTools.E_ALIGNMENT.RIGHT)); 

_concat.addContent
	('T'); 

_concat.addContent
	(KOSTAL_AF2024_Core_StringTools.F_FormatMask_UTF8
			(	WORD_TO_STRING(_ITime.TimeStruct.Hour), 
				'00', KOSTAL_AF2024_Core_StringTools.E_ALIGNMENT.RIGHT)); 

_concat.addContent
	(':'); 

_concat.addContent
	(KOSTAL_AF2024_Core_StringTools.F_FormatMask_UTF8
			(	WORD_TO_STRING(_ITime.TimeStruct.Minute), 
				'00', KOSTAL_AF2024_Core_StringTools.E_ALIGNMENT.RIGHT)); 

_concat.addContent
	(':'); 

_concat.addContent
	(KOSTAL_AF2024_Core_StringTools.F_FormatMask_UTF8
			(	WORD_TO_STRING(_ITime.TimeStruct.Second), 
				'00', KOSTAL_AF2024_Core_StringTools.E_ALIGNMENT.RIGHT)); 

GetTimeStamp:= _concat.getResult();

_concat.clear();
END_METHOD

METHOD PUBLIC linkConfig
VAR_INPUT
	CFG	:	I_T_CFG;
END_VAR

IF CFG = 0 THEN RETURN;	END_IF

IF NOT CFG.Valid THEN RETURN;	END_IF

IF CFG.HostName <> ''	THEN _HostName:= CFG.HostName;	END_IF
IF CFG.HostPort <> 0	THEN _HostPort:= CFG.HostPort;	END_IF

IF CFG.ClientName <> ''			THEN _ClientName:= CFG.ClientName;	END_IF
IF CFG.ClientProcess <> ''	THEN _ClientProcess:= CFG.ClientProcess;	END_IF
END_METHOD

METHOD PUBLIC LinkTime
VAR_INPUT
	Link	: KOSTAL_AF2024_Core_GetSystemTime.I_TimeSource;
END_VAR

IF Link <> 0 THEN	_ITime:= Link;	END_IF
END_METHOD

METHOD PUBLIC RedirectClient
VAR_INPUT
END_VAR

_clientRedirect:= TRUE;
END_METHOD

(*
Set Verbose level with target data
===================================
*)
METHOD PUBLIC Verbose

VAR_INPUT
	PathName	: KOSTAL_AF2024_Core_Settings.T_MaxString_UTF8;	
	FileName	: KOSTAL_AF2024_Core_Settings.T_MaxString_UTF8;
	Verbose		: E_Verbose;
END_VAR


IF Tc2_Standard.RIGHT(PathName, 1) = '\' THEN

	_Path_Logger:= PathName;	

ELSE

	_concat.clear();
	_concat.addContent(PathName);
	_concat.addContent('\');
	_Path_Logger:= _concat.getResult();
	_concat.clear();
	
END_IF

_File_Logger:= FileName;

_Verbose:= Verbose;
END_METHOD

METHOD PROTECTED _FBmain
VAR_INPUT
END_VAR


_deviceDefine();

IF NOT _isInit 																										THEN	_step.init();
ELSIF _THIS_CALLED <> _THIS_IN_PROCESS														THEN	_step.init();	
//ELSIF NOT _client.bConfigured AND _step.actual <> _ADDRESS_READY 	THEN	_step.init();
END_IF

_step.Header();

_isInit:= TRUE;
END_METHOD

END_FUNCTION_BLOCK

// Project Information/F_GetVersion
// This function has been automatically generated from the project information.
{attribute 'signature_flag' := '1073741824'}
{attribute 'TcGenerated'}
{attribute 'no-analysis'}
FUNCTION F_GetVersion : ST_LibVersion
VAR_INPUT
	
END_VAR

F_GetVersion.iMajor := 1;
F_GetVersion.iMinor := 0;
F_GetVersion.iBuild := 0;
F_GetVersion.iRevision := 0;
F_GetVersion.sVersion := '1.0.0.0';
F_GetVersion.nFlags := 1;

END_FUNCTION

// Project Information/F_GetTitle
// This function has been automatically generated from the project information.
{attribute 'signature_flag' := '1073741824'}
{attribute 'TcGenerated'}
{attribute 'no-analysis'}
FUNCTION F_GetTitle : WSTRING
VAR_INPUT
	
END_VAR

F_GetTitle := "KOSTAL.AF2024.Connectivity.LC";

END_FUNCTION

// 3_DUT/OptionalFlags/I_T_OptionalFlags
INTERFACE I_T_OptionalFlags EXTENDS _I_T_Copy

METHOD PUBLIC FlagsInRange : BOOL
VAR_INPUT
	FlagNumber	: UINT;	//1..
END_VAR
END_METHOD

METHOD PUBLIC get : BOOL
VAR_INPUT
	FlagNumber	: UINT;
END_VAR
END_METHOD

END_INTERFACE

// 3_DUT/OptionalFlags/I_T_OptionalFlags_Owner
INTERFACE I_T_OptionalFlags_Owner EXTENDS _I_T_Copy_Owner

METHOD PUBLIC clear
VAR_INPUT
END_VAR
END_METHOD

METHOD PUBLIC FlagsInRange : BOOL
VAR_INPUT
	FlagNumber	: UINT;	//1..
END_VAR
END_METHOD

METHOD PUBLIC get : BOOL
VAR_INPUT
	FlagNumber	: UINT;
END_VAR
END_METHOD

(*
	Return TRUE if Number has a valid Value
*)
METHOD PUBLIC set : BOOL
VAR_INPUT
	Number	: UINT;	//1..
	state	: BOOL;
END_VAR
END_METHOD

END_INTERFACE

// 3_DUT/OptionalFlags/T_OptionalFlags
FUNCTION_BLOCK PUBLIC T_OptionalFlags EXTENDS _T_Copy IMPLEMENTS I_T_OptionalFlags_Owner, I_T_OptionalFlags

VAR
	_optionalFlags		: ARRAY[1..SETTINGS.OPTIONAL_FLAGS_MAX] OF BOOL;
END_VAR

METHOD PUBLIC clear
VAR_INPUT
END_VAR

VAR
	_i: UINT;
END_VAR


FOR _i:= 1 TO SETTINGS.OPTIONAL_FLAGS_MAX DO
	_optionalFlags[_i]:= FALSE;
END_FOR
END_METHOD

METHOD PUBLIC CopyFrom : BOOL
VAR_INPUT
	IN	: KOSTAL_AF2024_Core_System.I_Interface;
END_VAR

VAR
	_IN		: I_T_OptionalFlags;
	_IN2	: I_T_OptionalFlags_Owner;
	_ui	: UINT;
END_VAR

IF NOT SUPER^.CopyFrom(IN) THEN 	;

ELSIF __QUERYINTERFACE(IN, _IN2) AND_THEN _IN2 <> 0 THEN 

	FOR _ui:= 1 TO SETTINGS.OPTIONAL_FLAGS_MAX DO
	
		_optionalFlags[_ui]:= _IN2.get(_ui);	
	
	END_FOR

	CopyFrom:= TRUE;
	
ELSIF __QUERYINTERFACE(IN, _IN) AND_THEN _IN <> 0 THEN 

	FOR _ui:= 1 TO SETTINGS.OPTIONAL_FLAGS_MAX DO
	
		_optionalFlags[_ui]:= _IN.get(_ui);	
	
	END_FOR

	CopyFrom:= TRUE;

END_IF
END_METHOD

METHOD PUBLIC FlagsInRange : BOOL
VAR_INPUT
	FlagNumber	: UINT;	//1..
END_VAR

FlagsInRange:= (FlagNumber >= 1) AND (FlagNumber <= SETTINGS.OPTIONAL_FLAGS_MAX);
END_METHOD

METHOD PUBLIC get : BOOL
VAR_INPUT
	FlagNumber	: UINT;
END_VAR

IF FlagsInRange(FlagNumber) THEN
	get:= _optionalFlags[FlagNumber];
ELSE
	get:= FALSE;
END_IF
END_METHOD

(*
	Return TRUE if Number has a valid Value
*)
METHOD PUBLIC set : BOOL
VAR_INPUT
	Number	: UINT;	//1..
	state	: BOOL;
END_VAR


IF FlagsInRange(Number) THEN
	_optionalFlags[Number]:= state;
	set:= TRUE;
ELSE
	set:= FALSE;
END_IF
END_METHOD

END_FUNCTION_BLOCK

// 3_DUT/OptionalStrings/I_T_OptionalStrings
INTERFACE I_T_OptionalStrings EXTENDS _I_T_Copy

METHOD PUBLIC get : KOSTAL_AF2024_Core_Settings.T_MaxString_UTF8
VAR_INPUT
	StringNumber	: UINT;
END_VAR
END_METHOD

METHOD PUBLIC StringsInRange : BOOL
VAR_INPUT
	Number	: UINT;	//1..
END_VAR
END_METHOD

END_INTERFACE

// 3_DUT/OptionalStrings/I_T_OptionalStrings_Owner
INTERFACE I_T_OptionalStrings_Owner EXTENDS _I_T_Copy_Owner

METHOD PUBLIC clear
VAR_INPUT
END_VAR
END_METHOD

METHOD PUBLIC get : KOSTAL_AF2024_Core_Settings.T_MaxString_UTF8
VAR_INPUT
	StringNumber	: UINT;
END_VAR
END_METHOD

(*
	Return TRUE if StringNumber has a valid Value
*)
METHOD PUBLIC set : BOOL
VAR_INPUT
	Number	: UINT;	//1..
	content	: KOSTAL_AF2024_Core_Settings.T_MaxString_UTF8;
END_VAR
END_METHOD

METHOD PUBLIC StringsInRange : BOOL
VAR_INPUT
	Number	: UINT;	//1..
END_VAR
END_METHOD

END_INTERFACE

// 3_DUT/OptionalStrings/T_OptionalStrings
FUNCTION_BLOCK PUBLIC T_OptionalStrings EXTENDS _T_Copy IMPLEMENTS I_T_OptionalStrings_Owner, I_T_OptionalStrings

VAR
	_optionalStrings	: ARRAY[1..SETTINGS.OPTIONAL_STRINGS_MAX] OF KOSTAL_AF2024_Core_Settings.T_MaxString_UTF8;
END_VAR

METHOD PUBLIC clear
VAR_INPUT
END_VAR

VAR
	_i: UINT;
END_VAR


FOR _i:= 1 TO SETTINGS.OPTIONAL_STRINGS_MAX DO
	_optionalStrings[_i]:= '';
END_FOR
END_METHOD

METHOD PUBLIC CopyFrom : BOOL
VAR_INPUT
	IN	: KOSTAL_AF2024_Core_System.I_Interface;
END_VAR

VAR
	_IN		: I_T_OptionalStrings;
	_IN2	: I_T_OptionalStrings_Owner;
	_ui		: UINT;
END_VAR

IF NOT SUPER^.CopyFrom(IN) THEN 	;

ELSIF __QUERYINTERFACE(IN, _IN2) AND_THEN _IN2 <> 0 THEN 

	FOR _ui:= 1 TO SETTINGS.OPTIONAL_STRINGS_MAX DO
	
		_optionalStrings[_ui]:= _IN2.get(_ui);	
	
	END_FOR

	CopyFrom:= TRUE;
	
ELSIF __QUERYINTERFACE(IN, _IN) AND_THEN _IN <> 0 THEN 
	
	FOR _ui:= 1 TO SETTINGS.OPTIONAL_STRINGS_MAX DO
	
		_optionalStrings[_ui]:= _IN.get(_ui);	
	
	END_FOR

	CopyFrom:= TRUE;

END_IF
END_METHOD

METHOD PUBLIC get : KOSTAL_AF2024_Core_Settings.T_MaxString_UTF8
VAR_INPUT
	StringNumber	: UINT;
END_VAR

IF StringsInRange(StringNumber) THEN
	get:= _optionalStrings[StringNumber];
ELSE
	get:= '';
END_IF
END_METHOD

(*
	Return TRUE if StringNumber has a valid Value
*)
METHOD PUBLIC set : BOOL
VAR_INPUT
	Number	: UINT;	//1..
	content	: KOSTAL_AF2024_Core_Settings.T_MaxString_UTF8;
END_VAR


IF StringsInRange(Number) THEN
	_optionalStrings[Number]:= content;
	set:= TRUE;
ELSE
	set:= FALSE;
END_IF
END_METHOD

METHOD PUBLIC StringsInRange : BOOL
VAR_INPUT
	Number	: UINT;	//1..
END_VAR

StringsInRange:= (Number >= 1) AND (Number <= SETTINGS.OPTIONAL_STRINGS_MAX);
END_METHOD

END_FUNCTION_BLOCK

// 3_DUT/PreviousProcess/ListOf/FB_ListOfPreviousProcess
FUNCTION_BLOCK FB_ListOfPreviousProcess  EXTENDS KOSTAL_AF2024_Core_ListOf._FB_Object_Base IMPLEMENTS I_ListOfPreviousProcess, I_ListOfPreviousProcess_CopyFrom, I_ListOfPreviousProcess_Owner

VAR
	_Dummy	: T_PreviousProcess;
END_VAR

(*
	Returns the typed interface in the reference variable.
	In the event of an error, the return value becomes FALSE and the interface refers to the {_Dummy}.
*)
METHOD PROTECTED _get_I : I_T_PreviousProcess

VAR_INPUT
	Member		: KOSTAL_AF2024_Core_System.I_Interface;
	rValid		: REFERENCE TO BOOL;
	Response	: KOSTAL_AF2024_Core_functionResponse.I_T_functionResponse_Owner;
END_VAR

VAR
	_iObj			: I_T_PreviousProcess;
END_VAR
//preset
_get_I:= _Dummy;
IF __ISVALIDREF(rValid)	THEN	rValid:= FALSE;	END_IF	

IF NOT _verifyMember(Member, Response)	THEN RETURN;	END_IF

//return dummy if no valid DUT is found
IF NOT __QUERYINTERFACE(Member, _iObj) OR_ELSE (_iObj = 0)	THEN		
	_setResultFail(Response, "__QueryInterface failed - return Dummy");	RETURN;	
END_IF

IF __ISVALIDREF(rValid)	THEN	rValid:= TRUE;	END_IF	
_setResultPass(Response, "Successful");

_get_I:= _iObj;
END_METHOD

(*
	Returns the typed owner interface in the reference variable.
	In the event of an error, the return value becomes FALSE and the interface refers to the {_Dummy}.
*)
METHOD PROTECTED _get_I_Owner : I_T_PreviousProcess_Owner

VAR_INPUT
	Member		: KOSTAL_AF2024_Core_System.I_Interface;
	rValid		: REFERENCE TO BOOL;
	Response	: KOSTAL_AF2024_Core_functionResponse.I_T_functionResponse_Owner;
END_VAR

VAR
	_iObj			: I_T_PreviousProcess_Owner;
END_VAR
//preset
_get_I_Owner:= _Dummy;

IF 		__ISVALIDREF(rValid)	THEN	rValid:= FALSE;	END_IF	

IF NOT _verifyMember(Member, Response)	THEN RETURN;	END_IF

//return dummy if no valid DUT is found
IF NOT __QUERYINTERFACE(Member, _iObj) OR_ELSE (_iObj = 0)	THEN	
	_setResultFail(Response, "__QueryInterface failed - return Dummy");	RETURN;	
END_IF

IF __ISVALIDREF(rValid)	THEN	rValid:= TRUE;	END_IF
_setResultPass(Response, "Successful");
_get_I_Owner:= _iObj;
END_METHOD

(*
	Cleans the custom class {FB_DUT} and removes it from memory.
*)
METHOD PROTECTED  _removePayLoad : BOOL
VAR_INPUT
	Member	: KOSTAL_AF2024_Core_System.I_Interface;
	Result	: KOSTAL_AF2024_Core_functionResponse.I_T_functionResponse_Owner;
END_VAR

VAR
	_iObj			: I_T_PreviousProcess_Owner;
	_pFB_DUT	:	POINTER TO T_PreviousProcess;
	_Success	: BOOL;
END_VAR


IF NOT SUPER^._removePayload(Member, Result)	THEN RETURN;	END_IF

_Success:= __QUERYINTERFACE(Member, _iObj);

IF NOT _Success	THEN	RETURN;	END_IF
IF _iObj = 0		THEN	RETURN;	END_IF

_iObj.Clear();

_Success  := __QUERYPOINTER(_iObj, _pFB_DUT);

IF NOT _Success	THEN	RETURN;	END_IF
IF _pFB_DUT = 0	THEN	RETURN;	END_IF

__DELETE(_pFB_DUT);
END_METHOD

(*
	Overload the method from the base class to verify the custom interface. 
	The local method {_get_I_Owner()} is used for this.
*)
METHOD PROTECTED _verifyMember : BOOL

VAR_INPUT
	Member	: KOSTAL_AF2024_Core_System.I_Interface;
	Result	: KOSTAL_AF2024_Core_functionResponse.I_T_functionResponse_Owner;
END_VAR

VAR
	_pObj	: POINTER TO T_PreviousProcess;
	_Success: BOOL;
END_VAR

IF NOT SUPER^._verifyMember(Member, Result)	THEN RETURN;	END_IF

_Success:= __QUERYPOINTER(Member, _pObj);

//return dummy if no valid Pointer to DUT is found
IF NOT _Success OR_ELSE (_pObj = 0)	THEN	_setResultFail(Result, "__QueryPointer failed");	RETURN; END_IF

_verifyMember:= TRUE;
END_METHOD

(*
	Add a new instance of FB_Dut and copy content from [IN] to the new instance
*)
METHOD PUBLIC Add_DUT : BOOL
VAR_INPUT
	IN				: KOSTAL_AF2024_Core_System.I_Interface;
	Response	: KOSTAL_AF2024_Core_functionResponse.I_T_functionResponse_Owner;
END_VAR

VAR
	_IN1	: I_T_PreviousProcess;
	_IN2	: I_T_PreviousProcess_Owner;
	_pDUT	: POINTER TO T_PreviousProcess;
END_VAR

IF IN = 0 THEN	RETURN;	END_IF


IF __QUERYINTERFACE(IN, _IN1) AND_THEN (_IN1 <> 0)	THEN


	_pDUT:= __NEW(T_PreviousProcess);
	
	IF _pDUT = 0 THEN	_setResultFail(Response, "cannot create new object"); RETURN; END_IF
	
	_pDUT^.CopyFrom(_IN1);
	
	Add_DUT:= _addMember(_pDUT^, Response);


ELSIF __QUERYINTERFACE(IN, _IN2) AND_THEN (_IN2 <> 0)	THEN


	_pDUT:= __NEW(T_PreviousProcess);
	
	IF _pDUT = 0 THEN	_setResultFail(Response, "cannot create new object"); RETURN; END_IF
	
	_pDUT^.CopyFrom(_IN2);
	
	Add_DUT:= _addMember(_pDUT^, Response);


END_IF
END_METHOD

(*
	Makes the protected method public.
*)
METHOD Clear

_clear();
END_METHOD

(*
	Copies the contents of another list {IN} into its own memory.
*)
METHOD PUBLIC CopyFrom
VAR_INPUT
	IN	: KOSTAL_AF2024_Core_System.I_Interface;
END_VAR

VAR
	_udi	: UDINT;

	_IN		: I_ListOfPreviousProcess;
	_IN_O	: I_ListOfPreviousProcess_Owner;

END_VAR

IF IN = 0 THEN RETURN;	END_IF

IF __QUERYINTERFACE(IN, _IN_O) AND_THEN _IN_O <> 0	THEN

	_clear();
	
	FOR _udi:= 1 TO _IN_O.NumberOfMember DO
		Add_DUT(_IN_O.Get_I_Owner(_udi, 0, 0), 0);
	END_FOR
	
ELSIF __QUERYINTERFACE(IN, _IN) AND_THEN _IN <> 0	THEN	

	_clear();
	
	FOR _udi:= 1 TO _IN.NumberOfMember DO
		Add_DUT(_IN.Get_I(_udi, 0, 0), 0);
	END_FOR

END_IF
END_METHOD

(*
	Copies the own content into another list created at the parameter {IN}.
*)
METHOD PUBLIC CopyTo
VAR_INPUT
	IN	: KOSTAL_AF2024_Core_System.I_Interface;
END_VAR

VAR
	_IN	: I_ListOfPreviousProcess_CopyFrom;
END_VAR

IF (IN = 0) OR_ELSE NOT __QUERYINTERFACE(IN, _IN) OR_ELSE (_IN = 0) THEN	RETURN;	END_IF

_IN.CopyFrom(THIS^);
END_METHOD

(*
	Deletes the class specified with the {Number} from the list.
*)
METHOD PUBLIC Delete_DUT : BOOL
VAR_INPUT
	Number		: UDINT;	//Number of DUT in List
	Response	: KOSTAL_AF2024_Core_functionResponse.I_T_functionResponse_Owner;
END_VAR

VAR
	//_response	: KOSTAL_AF2024_Core_functionResponse.T_functionResponse;
	_Success	: BOOL;
	_Member		: KOSTAL_AF2024_Core_System.I_Interface;
END_VAR

IF Number = 0 THEN	_setResultFail(Response, "Number is out of range (1..n)"); RETURN; END_IF

Delete_DUT:= _removeMemberByIndex(Number - 1, Response);
END_METHOD

(*
	Get readonly access to content of Member with {Number}
*) 
METHOD Get_I : I_T_PreviousProcess

VAR_INPUT
	Number		: UDINT;
	rValid		: REFERENCE TO BOOL;
	Response	: KOSTAL_AF2024_Core_functionResponse.I_T_functionResponse_Owner;
END_VAR

VAR
	_Member	: KOSTAL_AF2024_Core_System.I_Interface;
END_VAR

//preset
Get_I:=	_Dummy; 
IF __ISVALIDREF(rValid)	THEN	rValid:= FALSE;	END_IF	

IF Number = 0 THEN _setResultFail(Response, "Number is out of range (1..n)"); RETURN; END_IF

IF _findMemberByIndex(Number - 1, _Member, Response) THEN
	Get_I:= _get_I(_Member, rValid, Response);
END_IF
END_METHOD

METHOD PUBLIC Get_I_ByProcessName : I_T_PreviousProcess

VAR_INPUT
	ProcessName	: KOSTAL_AF2024_Core_Settings.T_MaxString_UTF8;
	rValid			: REFERENCE TO BOOL;
	Response		: KOSTAL_AF2024_Core_functionResponse.I_T_functionResponse_Owner;
END_VAR

VAR
	_udi		: UDINT;
	_obj		: I_T_PreviousProcess;
END_VAR
//preset
Get_I_ByProcessName:= _Dummy;

IF __ISVALIDREF(rValid) THEN rValid:= FALSE;	END_IF

FOR _udi:= 1 TO _NumberOfMember DO
	
	_obj:= Get_I(_udi, rValid, Response);		

	IF _obj.processName = ProcessName THEN	Get_I_ByProcessName:= _obj;	RETURN;	END_IF

END_FOR

IF __ISVALIDREF(rValid) THEN rValid:= FALSE;	END_IF
_setResultFail(Response, "no entry with this ID found");
END_METHOD

(*
	Get full access to content of Member with {Number}
*) 
METHOD Get_I_Owner : I_T_PreviousProcess_Owner

VAR_INPUT
	Number		: UDINT;
	rValid		: REFERENCE TO BOOL;
	Response	: KOSTAL_AF2024_Core_functionResponse.I_T_functionResponse_Owner;
END_VAR

VAR
	_Member	: KOSTAL_AF2024_Core_System.I_Interface;
END_VAR
//preset

Get_I_Owner:= _Dummy;

IF __ISVALIDREF(rValid)	THEN	rValid:= FALSE;	END_IF	

IF Number = 0 THEN _setResultFail(Response, "Number is out of range (1..n)"); RETURN; END_IF

IF _findMemberByIndex(Number - 1, _Member, Response) THEN
	Get_I_Owner:= _get_I_Owner(_Member, rValid, Response);
END_IF
END_METHOD

(*
	Number of Member in list.
*)
PROPERTY NumberOfMember : UDINT
GET

NumberOfMember:= SUPER^._NumberOfMember;
END_GET
END_PROPERTY

END_FUNCTION_BLOCK

// 3_DUT/PreviousProcess/ListOf/I_ListOfPreviousProcess
INTERFACE I_ListOfPreviousProcess EXTENDS KOSTAL_AF2024_Core_ListOf._I_Object_Base

(*
	Copies the own content into another list created at the parameter {IN}.
*)
METHOD PUBLIC CopyTo
VAR_INPUT
	IN	: KOSTAL_AF2024_Core_System.I_Interface;
END_VAR
END_METHOD

(*
	Get readonly access to content of Member with {Number}
*) 
METHOD Get_I : I_T_PreviousProcess

VAR_INPUT
	Number		: UDINT;
	rValid		: REFERENCE TO BOOL;
	Response	: KOSTAL_AF2024_Core_functionResponse.I_T_functionResponse_Owner;
END_VAR
END_METHOD

METHOD PUBLIC Get_I_ByProcessName : I_T_PreviousProcess

VAR_INPUT
	ProcessName	: KOSTAL_AF2024_Core_Settings.T_MaxString_UTF8;
	rValid			: REFERENCE TO BOOL;
	Response		: KOSTAL_AF2024_Core_functionResponse.I_T_functionResponse_Owner;
END_VAR
END_METHOD

(*
	Number of Member in list.
*)
PROPERTY NumberOfMember : UDINT
GET
END_GET
END_PROPERTY

END_INTERFACE

// 3_DUT/PreviousProcess/I_T_PreviousProcess
INTERFACE I_T_PreviousProcess EXTENDS _I_T_Copy

PROPERTY PUBLIC articlenumberRegex : KOSTAL_AF2024_Core_Settings.T_MaxString_UTF8
GET
END_GET
END_PROPERTY

PROPERTY PUBLIC databaseName : KOSTAL_AF2024_Core_Settings.T_MaxString_UTF8
GET
END_GET
END_PROPERTY

PROPERTY PUBLIC PreviousProcesses : KOSTAL_AF2024_Core_ListOf.I_ListOfString_UTF8
GET
END_GET
END_PROPERTY

PROPERTY PUBLIC processName : KOSTAL_AF2024_Core_Settings.T_MaxString_UTF8
GET
END_GET
END_PROPERTY

PROPERTY PUBLIC processStamp : KOSTAL_AF2024_Core_Settings.T_MaxString_UTF8
GET
END_GET
END_PROPERTY

PROPERTY PUBLIC searchMode : DINT
GET
END_GET
END_PROPERTY

PROPERTY PUBLIC useOnlyTable : KOSTAL_AF2024_Core_Settings.T_MaxString_UTF8
GET
END_GET
END_PROPERTY

END_INTERFACE

// 3_DUT/PreviousProcess/ListOf/I_ListOfPreviousProcess_CopyFrom
INTERFACE I_ListOfPreviousProcess_CopyFrom EXTENDS KOSTAL_AF2024_Core_System.I_Interface

METHOD PUBLIC CopyFrom
VAR_INPUT
	IN	: KOSTAL_AF2024_Core_System.I_Interface;
END_VAR
END_METHOD

END_INTERFACE

// 3_DUT/PreviousProcess/ListOf/I_ListOfPreviousProcess_Owner
INTERFACE I_ListOfPreviousProcess_Owner EXTENDS KOSTAL_AF2024_Core_ListOf._I_Object_Base_Owner

(*
	Add a new instance of FB_Dut and copy content from [IN] to the new instance
*)
METHOD PUBLIC Add_DUT : BOOL
VAR_INPUT
	IN				: KOSTAL_AF2024_Core_System.I_Interface;
	Response	: KOSTAL_AF2024_Core_functionResponse.I_T_functionResponse_Owner;
END_VAR
END_METHOD

(*
	Makes the protected method public.
*)
METHOD Clear
END_METHOD

(*
	Copies the contents of another list {IN} into its own memory.
*)
METHOD PUBLIC CopyFrom
VAR_INPUT
	IN	: KOSTAL_AF2024_Core_System.I_Interface;
END_VAR
END_METHOD

(*
	Copies the own content into another list created at the parameter {IN}.
*)
METHOD PUBLIC CopyTo
VAR_INPUT
	IN	: KOSTAL_AF2024_Core_System.I_Interface;
END_VAR
END_METHOD

(*
	Deletes the class specified with the {Number} from the list.
*)
METHOD PUBLIC Delete_DUT : BOOL
VAR_INPUT
	Number		: UDINT;	//Number of DUT in List
	Response	: KOSTAL_AF2024_Core_functionResponse.I_T_functionResponse_Owner;
END_VAR
END_METHOD

(*
	Get readonly access to content of Member with {Number}
*) 
METHOD Get_I : I_T_PreviousProcess

VAR_INPUT
	Number		: UDINT;
	rValid		: REFERENCE TO BOOL;
	Response	: KOSTAL_AF2024_Core_functionResponse.I_T_functionResponse_Owner;
END_VAR
END_METHOD

METHOD PUBLIC Get_I_ByProcessName : I_T_PreviousProcess

VAR_INPUT
	ProcessName	: KOSTAL_AF2024_Core_Settings.T_MaxString_UTF8;
	rValid			: REFERENCE TO BOOL;
	Response		: KOSTAL_AF2024_Core_functionResponse.I_T_functionResponse_Owner;
END_VAR
END_METHOD

(*
	Get full access to content of Member with {Number}
*) 
METHOD Get_I_Owner : I_T_PreviousProcess_Owner

VAR_INPUT
	Number		: UDINT;
	rValid		: REFERENCE TO BOOL;
	Response	: KOSTAL_AF2024_Core_functionResponse.I_T_functionResponse_Owner;
END_VAR
END_METHOD

(*
	Number of Member in list.
*)
PROPERTY NumberOfMember : UDINT
GET
END_GET
END_PROPERTY

END_INTERFACE

// 3_DUT/PreviousProcess/I_T_PreviousProcess_Owner
INTERFACE I_T_PreviousProcess_Owner EXTENDS _I_T_Copy_Owner

PROPERTY PUBLIC articlenumberRegex : KOSTAL_AF2024_Core_Settings.T_MaxString_UTF8
GET
END_GET
SET
END_SET
END_PROPERTY

METHOD PUBLIC clear
VAR_INPUT
END_VAR
END_METHOD

PROPERTY PUBLIC databaseName : KOSTAL_AF2024_Core_Settings.T_MaxString_UTF8
GET
END_GET
SET
END_SET
END_PROPERTY

PROPERTY PUBLIC PreviousProcesses_Owner : KOSTAL_AF2024_Core_ListOf.I_ListOfString_UTF8_Owner
GET
END_GET
END_PROPERTY

PROPERTY PUBLIC processName : KOSTAL_AF2024_Core_Settings.T_MaxString_UTF8
GET
END_GET
SET
END_SET
END_PROPERTY

PROPERTY PUBLIC processStamp : KOSTAL_AF2024_Core_Settings.T_MaxString_UTF8
GET
END_GET
SET
END_SET
END_PROPERTY

PROPERTY PUBLIC searchMode : DINT
GET
END_GET
SET
END_SET
END_PROPERTY

PROPERTY PUBLIC useOnlyTable : KOSTAL_AF2024_Core_Settings.T_MaxString_UTF8
GET
END_GET
SET
END_SET
END_PROPERTY

END_INTERFACE

// 3_DUT/PreviousProcess/T_PreviousProcess
{attribute 'enable_dynamic_creation'}
FUNCTION_BLOCK PUBLIC T_PreviousProcess EXTENDS _T_Copy IMPLEMENTS I_T_PreviousProcess_Owner, I_T_PreviousProcess

VAR
  _processName				: KOSTAL_AF2024_Core_Settings.T_MaxString_UTF8;	//": "^[0-9]{8}-(([0-9]{2})|([0-9]{4}))$",
  _processStamp				: KOSTAL_AF2024_Core_Settings.T_MaxString_UTF8;	//": "^([A-Z0-9]{13})$|^([0-9]{14})$",
  _databaseName				: KOSTAL_AF2024_Core_Settings.T_MaxString_UTF8;	//": test,
	_useOnlyTable				: KOSTAL_AF2024_Core_Settings.T_MaxString_UTF8;	//": lc_test,
	_searchMode					: DINT;	//": 0
  _articlenumberRegex	: KOSTAL_AF2024_Core_Settings.T_MaxString_UTF8;	//": "^[0-9]{8}-(([0-9]{2})|([0-9]{4}))$",
	_previousProcesses	: KOSTAL_AF2024_Core_ListOf.FB_ListOfString_UTF8;
END_VAR

PROPERTY PUBLIC articlenumberRegex : KOSTAL_AF2024_Core_Settings.T_MaxString_UTF8
GET

articlenumberRegex	:= _articlenumberRegex;
END_GET
SET

_articlenumberRegex	:= articlenumberRegex;
END_SET
END_PROPERTY

METHOD PUBLIC clear
VAR_INPUT
END_VAR

_processName				:= '';
_processStamp				:= '';
_databaseName				:= '';
_useOnlyTable				:= '';
_searchMode					:= 0;
_articlenumberRegex	:= '';

_previousProcesses.clear();
END_METHOD

METHOD PUBLIC CopyFrom : BOOL
VAR_INPUT
	IN	: KOSTAL_AF2024_Core_System.I_Interface;
END_VAR

VAR
	_IN	: I_T_PreviousProcess;
	_ui	: UDINT;
END_VAR

IF NOT SUPER^.CopyFrom(IN) THEN RETURN;	END_IF

IF NOT __QUERYINTERFACE(IN, _IN) OR_ELSE _IN = 0 THEN RETURN;	END_IF

_processName				:= _IN.processName;
_processStamp				:= _IN.processStamp;
_databaseName				:= _IN.databaseName;
_useOnlyTable				:= _IN.useOnlyTable;
_searchMode					:= _IN.searchMode;
_articlenumberRegex	:= _IN.articlenumberRegex;

_previousProcesses.clear();

FOR _ui:= 1 TO _IN.PreviousProcesses.NumberOfLines DO
	_previousProcesses.addLine(_IN.PreviousProcesses.line_GET(_ui));
END_FOR 

CopyFrom:= TRUE;
END_METHOD

PROPERTY PUBLIC databaseName : KOSTAL_AF2024_Core_Settings.T_MaxString_UTF8
GET

databaseName:= _databaseName;
END_GET
SET

_databaseName:= databaseName;
END_SET
END_PROPERTY

PROPERTY PUBLIC PreviousProcesses : KOSTAL_AF2024_Core_ListOf.I_ListOfString_UTF8
GET

PreviousProcesses:= _previousProcesses;
END_GET
END_PROPERTY

PROPERTY PUBLIC PreviousProcesses_Owner : KOSTAL_AF2024_Core_ListOf.I_ListOfString_UTF8_Owner
GET

PreviousProcesses_Owner := _previousProcesses;
END_GET
END_PROPERTY

PROPERTY PUBLIC processName : KOSTAL_AF2024_Core_Settings.T_MaxString_UTF8
GET

processName:= _processName;
END_GET
SET

_processName:= processName;
END_SET
END_PROPERTY

PROPERTY PUBLIC processStamp : KOSTAL_AF2024_Core_Settings.T_MaxString_UTF8
GET

processStamp:= _processStamp;
END_GET
SET

_processStamp:= processStamp;
END_SET
END_PROPERTY

PROPERTY PUBLIC searchMode : DINT
GET

searchMode:= _searchMode;
END_GET
SET

_searchMode:= searchMode;
END_SET
END_PROPERTY

PROPERTY PUBLIC useOnlyTable : KOSTAL_AF2024_Core_Settings.T_MaxString_UTF8
GET

useOnlyTable:= _useOnlyTable;
END_GET
SET

_useOnlyTable:= useOnlyTable;
END_SET
END_PROPERTY

END_FUNCTION_BLOCK

// 3_DUT/ProcessConfig/ListOf/FB_ListOfProcessConfig
FUNCTION_BLOCK FB_ListOfProcessConfig  EXTENDS KOSTAL_AF2024_Core_ListOf._FB_Object_Base IMPLEMENTS I_ListOfProcessConfig, I_ListOfProcessConfig_CopyFrom, I_ListOfProcessConfig_Owner

VAR
	_Dummy	: T_ProcessConfig;
END_VAR

(*
	Returns the typed interface in the reference variable.
	In the event of an error, the return value becomes FALSE and the interface refers to the {_Dummy}.
*)
METHOD PROTECTED _get_I : I_T_ProcessConfig

VAR_INPUT
	Member		: KOSTAL_AF2024_Core_System.I_Interface;
	rValid		: REFERENCE TO BOOL;
	Response	: KOSTAL_AF2024_Core_functionResponse.I_T_functionResponse_Owner;
END_VAR

VAR
	_iObj			: I_T_ProcessConfig;
END_VAR
//preset
_get_I:= _Dummy;
IF __ISVALIDREF(rValid)	THEN	rValid:= FALSE;	END_IF	

IF NOT _verifyMember(Member, Response)	THEN RETURN;	END_IF

//return dummy if no valid DUT is found
IF NOT __QUERYINTERFACE(Member, _iObj) OR_ELSE (_iObj = 0)	THEN		
	_setResultFail(Response, "__QueryInterface failed - return Dummy");	RETURN;	
END_IF

IF __ISVALIDREF(rValid)	THEN	rValid:= TRUE;	END_IF	
_setResultPass(Response, "Successful");

_get_I:= _iObj;
END_METHOD

(*
	Returns the typed owner interface in the reference variable.
	In the event of an error, the return value becomes FALSE and the interface refers to the {_Dummy}.
*)
METHOD PROTECTED _get_I_Owner : I_T_ProcessConfig_Owner

VAR_INPUT
	Member		: KOSTAL_AF2024_Core_System.I_Interface;
	rValid		: REFERENCE TO BOOL;
	Response	: KOSTAL_AF2024_Core_functionResponse.I_T_functionResponse_Owner;
END_VAR

VAR
	_iObj			: I_T_ProcessConfig_Owner;
END_VAR
//preset
_get_I_Owner:= _Dummy;

IF 		__ISVALIDREF(rValid)	THEN	rValid:= FALSE;	END_IF	

IF NOT _verifyMember(Member, Response)	THEN RETURN;	END_IF

//return dummy if no valid DUT is found
IF NOT __QUERYINTERFACE(Member, _iObj) OR_ELSE (_iObj = 0)	THEN	
	_setResultFail(Response, "__QueryInterface failed - return Dummy");	RETURN;	
END_IF

IF __ISVALIDREF(rValid)	THEN	rValid:= TRUE;	END_IF
_setResultPass(Response, "Successful");
_get_I_Owner:= _iObj;
END_METHOD

(*
	Cleans the custom class {FB_DUT} and removes it from memory.
*)
METHOD PROTECTED  _removePayLoad : BOOL
VAR_INPUT
	Member	: KOSTAL_AF2024_Core_System.I_Interface;
	Result	: KOSTAL_AF2024_Core_functionResponse.I_T_functionResponse_Owner;
END_VAR

VAR
	_iObj			: I_T_ProcessConfig_Owner;
	_pFB_DUT	:	POINTER TO T_ProcessConfig;
	_Success	: BOOL;
END_VAR


IF NOT SUPER^._removePayload(Member, Result)	THEN RETURN;	END_IF

_Success:= __QUERYINTERFACE(Member, _iObj);

IF NOT _Success	THEN	RETURN;	END_IF
IF _iObj = 0		THEN	RETURN;	END_IF

_iObj.Clear();

_Success  := __QUERYPOINTER(_iObj, _pFB_DUT);

IF NOT _Success	THEN	RETURN;	END_IF
IF _pFB_DUT = 0	THEN	RETURN;	END_IF

__DELETE(_pFB_DUT);
END_METHOD

(*
	Overload the method from the base class to verify the custom interface. 
	The local method {_get_I_Owner()} is used for this.
*)
METHOD PROTECTED _verifyMember : BOOL

VAR_INPUT
	Member	: KOSTAL_AF2024_Core_System.I_Interface;
	Result	: KOSTAL_AF2024_Core_functionResponse.I_T_functionResponse_Owner;
END_VAR

VAR
	_pObj	: POINTER TO T_ProcessConfig;
	_Success: BOOL;
END_VAR

IF NOT SUPER^._verifyMember(Member, Result)	THEN RETURN;	END_IF

_Success:= __QUERYPOINTER(Member, _pObj);

//return dummy if no valid Pointer to DUT is found
IF NOT _Success OR_ELSE (_pObj = 0)	THEN	_setResultFail(Result, "__QueryPointer failed");	RETURN; END_IF

_verifyMember:= TRUE;
END_METHOD

(*
	Add a new instance of FB_Dut and copy content from [IN] to the new instance
*)
METHOD PUBLIC Add_DUT : BOOL
VAR_INPUT
	IN				: KOSTAL_AF2024_Core_System.I_Interface;
	Response	: KOSTAL_AF2024_Core_functionResponse.I_T_functionResponse_Owner;
END_VAR

VAR
	_IN1	: I_T_ProcessConfig;
	_IN2	: I_T_ProcessConfig_Owner;
	_pDUT	: POINTER TO T_ProcessConfig;
END_VAR

IF IN = 0 THEN	RETURN;	END_IF


IF __QUERYINTERFACE(IN, _IN1) AND_THEN (_IN1 <> 0)	THEN


	_pDUT:= __NEW(T_ProcessConfig);
	
	IF _pDUT = 0 THEN	_setResultFail(Response, "cannot create new object"); RETURN; END_IF
	
	_pDUT^.CopyFrom(_IN1);
	
	Add_DUT:= _addMember(_pDUT^, Response);


ELSIF __QUERYINTERFACE(IN, _IN2) AND_THEN (_IN2 <> 0)	THEN


	_pDUT:= __NEW(T_ProcessConfig);
	
	IF _pDUT = 0 THEN	_setResultFail(Response, "cannot create new object"); RETURN; END_IF
	
	_pDUT^.CopyFrom(_IN2);
	
	Add_DUT:= _addMember(_pDUT^, Response);


END_IF
END_METHOD

(*
	Makes the protected method public.
*)
METHOD Clear

_clear();
END_METHOD

(*
	Copies the contents of another list {IN} into its own memory.
*)
METHOD PUBLIC CopyFrom
VAR_INPUT
	IN	: KOSTAL_AF2024_Core_System.I_Interface;
END_VAR

VAR
	_udi	: UDINT;

	_IN		: I_ListOfProcessConfig;
	_IN_O	: I_ListOfProcessConfig_Owner;

END_VAR

IF IN = 0 THEN RETURN;	END_IF

IF __QUERYINTERFACE(IN, _IN_O) AND_THEN _IN_O <> 0	THEN

	_clear();
	
	FOR _udi:= 1 TO _IN_O.NumberOfMember DO
		Add_DUT(_IN_O.Get_I_Owner(_udi, 0, 0), 0);
	END_FOR
	
ELSIF __QUERYINTERFACE(IN, _IN) AND_THEN _IN <> 0	THEN	

	_clear();
	
	FOR _udi:= 1 TO _IN.NumberOfMember DO
		Add_DUT(_IN.Get_I(_udi, 0, 0), 0);
	END_FOR

END_IF
END_METHOD

(*
	Copies the own content into another list created at the parameter {IN}.
*)
METHOD PUBLIC CopyTo
VAR_INPUT
	IN	: KOSTAL_AF2024_Core_System.I_Interface;
END_VAR

VAR
	_IN	: I_ListOfPreviousProcess_CopyFrom;
END_VAR

IF (IN = 0) OR_ELSE NOT __QUERYINTERFACE(IN, _IN) OR_ELSE (_IN = 0) THEN	RETURN;	END_IF

_IN.CopyFrom(THIS^);
END_METHOD

(*
	Deletes the class specified with the {Number} from the list.
*)
METHOD PUBLIC Delete_DUT : BOOL
VAR_INPUT
	Number		: UDINT;	//Number of DUT in List
	Response	: KOSTAL_AF2024_Core_functionResponse.I_T_functionResponse_Owner;
END_VAR

VAR
	//_response	: KOSTAL_AF2024_Core_functionResponse.T_functionResponse;
	_Success	: BOOL;
	_Member		: KOSTAL_AF2024_Core_System.I_Interface;
END_VAR

IF Number = 0 THEN	_setResultFail(Response, "Number is out of range (1..n)"); RETURN; END_IF

Delete_DUT:= _removeMemberByIndex(Number - 1, Response);
END_METHOD

(*
	Get readonly access to content of Member with {Number}
*) 
METHOD Get_I : I_T_ProcessConfig

VAR_INPUT
	Number		: UDINT;
	rValid		: REFERENCE TO BOOL;
	Response	: KOSTAL_AF2024_Core_functionResponse.I_T_functionResponse_Owner;
END_VAR

VAR
	_Member	: KOSTAL_AF2024_Core_System.I_Interface;
END_VAR

//preset
Get_I:=	_Dummy; 
IF __ISVALIDREF(rValid)	THEN	rValid:= FALSE;	END_IF	

IF Number = 0 THEN _setResultFail(Response, "Number is out of range (1..n)"); RETURN; END_IF

IF _findMemberByIndex(Number - 1, _Member, Response) THEN
	Get_I:= _get_I(_Member, rValid, Response);
END_IF
END_METHOD

(*
	Get full access to content of Member with {Number}
*) 
METHOD Get_I_Owner : I_T_ProcessConfig_Owner

VAR_INPUT
	Number		: UDINT;
	rValid		: REFERENCE TO BOOL;
	Response	: KOSTAL_AF2024_Core_functionResponse.I_T_functionResponse_Owner;
END_VAR

VAR
	_Member	: KOSTAL_AF2024_Core_System.I_Interface;
END_VAR
//preset

Get_I_Owner:= _Dummy;

IF __ISVALIDREF(rValid)	THEN	rValid:= FALSE;	END_IF	

IF Number = 0 THEN _setResultFail(Response, "Number is out of range (1..n)"); RETURN; END_IF

IF _findMemberByIndex(Number - 1, _Member, Response) THEN
	Get_I_Owner:= _get_I_Owner(_Member, rValid, Response);
END_IF
END_METHOD

(*
	Number of Member in list.
*)
PROPERTY NumberOfMember : UDINT
GET

NumberOfMember:= SUPER^._NumberOfMember;
END_GET
END_PROPERTY

END_FUNCTION_BLOCK

// 3_DUT/ProcessConfig/ListOf/I_ListOfProcessConfig
INTERFACE I_ListOfProcessConfig EXTENDS KOSTAL_AF2024_Core_ListOf._I_Object_Base

(*
	Copies the own content into another list created at the parameter {IN}.
*)
METHOD PUBLIC CopyTo
VAR_INPUT
	IN	: KOSTAL_AF2024_Core_System.I_Interface;
END_VAR
END_METHOD

(*
	Get readonly access to content of Member with {Number}
*) 
METHOD Get_I : I_T_ProcessConfig

VAR_INPUT
	Number		: UDINT;
	rValid		: REFERENCE TO BOOL;
	Response	: KOSTAL_AF2024_Core_functionResponse.I_T_functionResponse_Owner;
END_VAR
END_METHOD

(*
	Number of Member in list.
*)
PROPERTY NumberOfMember : UDINT
GET
END_GET
END_PROPERTY

END_INTERFACE

// 3_DUT/ProcessConfig/I_T_ProcessConfig
INTERFACE I_T_ProcessConfig EXTENDS _I_T_Copy

PROPERTY PUBLIC activeCheckFQDN : BOOL
GET
END_GET
END_PROPERTY

PROPERTY PUBLIC allowedFQDN : KOSTAL_AF2024_Core_Settings.T_MaxString_UTF8
GET
END_GET
END_PROPERTY

PROPERTY PUBLIC articlenumberRegex : KOSTAL_AF2024_Core_Settings.T_MaxString_UTF8
GET
END_GET
END_PROPERTY

PROPERTY PUBLIC PreviousProcesses : I_ListOfPreviousProcess
GET
END_GET
END_PROPERTY

PROPERTY PUBLIC serialnumberRegex : KOSTAL_AF2024_Core_Settings.T_MaxString_UTF8
GET
END_GET
END_PROPERTY

PROPERTY PUBLIC traceID : DINT
GET
END_GET
END_PROPERTY

END_INTERFACE

// 3_DUT/ProcessConfig/ListOf/I_ListOfProcessConfig_CopyFrom
INTERFACE I_ListOfProcessConfig_CopyFrom EXTENDS KOSTAL_AF2024_Core_System.I_Interface

METHOD PUBLIC CopyFrom
VAR_INPUT
	IN	: KOSTAL_AF2024_Core_System.I_Interface;
END_VAR
END_METHOD

END_INTERFACE

// 3_DUT/ProcessConfig/ListOf/I_ListOfProcessConfig_Owner
INTERFACE I_ListOfProcessConfig_Owner EXTENDS KOSTAL_AF2024_Core_ListOf._I_Object_Base_Owner

(*
	Add a new instance of FB_Dut and copy content from [IN] to the new instance
*)
METHOD PUBLIC Add_DUT : BOOL
VAR_INPUT
	IN				: KOSTAL_AF2024_Core_System.I_Interface;
	Response	: KOSTAL_AF2024_Core_functionResponse.I_T_functionResponse_Owner;
END_VAR
END_METHOD

(*
	Makes the protected method public.
*)
METHOD Clear
END_METHOD

(*
	Copies the contents of another list {IN} into its own memory.
*)
METHOD PUBLIC CopyFrom
VAR_INPUT
	IN	: KOSTAL_AF2024_Core_System.I_Interface;
END_VAR
END_METHOD

(*
	Copies the own content into another list created at the parameter {IN}.
*)
METHOD PUBLIC CopyTo
VAR_INPUT
	IN	: KOSTAL_AF2024_Core_System.I_Interface;
END_VAR
END_METHOD

(*
	Deletes the class specified with the {Number} from the list.
*)
METHOD PUBLIC Delete_DUT : BOOL
VAR_INPUT
	Number		: UDINT;	//Number of DUT in List
	Response	: KOSTAL_AF2024_Core_functionResponse.I_T_functionResponse_Owner;
END_VAR
END_METHOD

(*
	Get readonly access to content of Member with {Number}
*) 
METHOD Get_I : I_T_ProcessConfig

VAR_INPUT
	Number		: UDINT;
	rValid		: REFERENCE TO BOOL;
	Response	: KOSTAL_AF2024_Core_functionResponse.I_T_functionResponse_Owner;
END_VAR
END_METHOD

(*
	Get full access to content of Member with {Number}
*) 
METHOD Get_I_Owner : I_T_ProcessConfig_Owner

VAR_INPUT
	Number		: UDINT;
	rValid		: REFERENCE TO BOOL;
	Response	: KOSTAL_AF2024_Core_functionResponse.I_T_functionResponse_Owner;
END_VAR
END_METHOD

(*
	Number of Member in list.
*)
PROPERTY NumberOfMember : UDINT
GET
END_GET
END_PROPERTY

END_INTERFACE

// 3_DUT/ProcessConfig/I_T_ProcessConfig_Owner
INTERFACE I_T_ProcessConfig_Owner EXTENDS _I_T_Copy_Owner

PROPERTY PUBLIC activeCheckFQDN : BOOL
GET
END_GET
SET
END_SET
END_PROPERTY

PROPERTY PUBLIC allowedFQDN : KOSTAL_AF2024_Core_Settings.T_MaxString_UTF8
GET
END_GET
SET
END_SET
END_PROPERTY

PROPERTY PUBLIC articlenumberRegex : KOSTAL_AF2024_Core_Settings.T_MaxString_UTF8
GET
END_GET
SET
END_SET
END_PROPERTY

METHOD PUBLIC clear
VAR_INPUT
END_VAR
END_METHOD

PROPERTY PUBLIC PreviousProcesses_Owner : I_ListOfPreviousProcess_Owner
GET
END_GET
END_PROPERTY

PROPERTY PUBLIC serialnumberRegex : KOSTAL_AF2024_Core_Settings.T_MaxString_UTF8
GET
END_GET
SET
END_SET
END_PROPERTY

PROPERTY PUBLIC traceID : DINT
GET
END_GET
SET
END_SET
END_PROPERTY

END_INTERFACE

// 3_DUT/ProcessConfig/T_ProcessConfig
{attribute 'enable_dynamic_creation'}
FUNCTION_BLOCK PUBLIC T_ProcessConfig EXTENDS _T_Copy IMPLEMENTS I_T_ProcessConfig_Owner, I_T_ProcessConfig

VAR
  _articlenumberRegex	: KOSTAL_AF2024_Core_Settings.T_MaxString_UTF8;	//": "^[0-9]{8}-(([0-9]{2})|([0-9]{4}))$",
  _serialnumberRegex	: KOSTAL_AF2024_Core_Settings.T_MaxString_UTF8;	//": "^([A-Z0-9]{13})$|^([0-9]{14})$",
  _traceID						: DINT;	//": 99056,
	_activeCheckFQDN		: BOOL;
	_allowedFQDN				: KOSTAL_AF2024_Core_Settings.T_MaxString_UTF8;
	_previousProcesses	: FB_ListOfPreviousProcess;
END_VAR

PROPERTY PUBLIC activeCheckFQDN : BOOL
GET

activeCheckFQDN:= _activeCheckFQDN;
END_GET
SET

_activeCheckFQDN:= activeCheckFQDN;
END_SET
END_PROPERTY

PROPERTY PUBLIC allowedFQDN : KOSTAL_AF2024_Core_Settings.T_MaxString_UTF8
GET

allowedFQDN:= _allowedFQDN;
END_GET
SET

_allowedFQDN:= allowedFQDN;
END_SET
END_PROPERTY

PROPERTY PUBLIC articlenumberRegex : KOSTAL_AF2024_Core_Settings.T_MaxString_UTF8
GET

articlenumberRegex	:= _articlenumberRegex;
END_GET
SET

_articlenumberRegex	:= articlenumberRegex;
END_SET
END_PROPERTY

METHOD PUBLIC clear
VAR_INPUT
END_VAR

